(* IEC 61131-3 sources: daoli-st-library/DL_Motion (part 21) *)

(* ---- FB_DL_ZoneSpeedTrim.st ---- *)
(*==============================================================================
 * 组件名称 (Component)  : FB_DL_ZoneSpeedTrim
 * 所属子库 (Sublibrary) : DL_Motion
 * 当前版本 (Version)    : 1.0.0
 * 兼容性   (Platform)   : CODESYS 3.5+ / TwinCAT 3 / 汇川 InoProShop / 施耐德 Machine Expert
 *                         仅依赖 Standard.library（MIN / MAX / ABS），零厂商私有库
 * 功能描述 (Function)   : 轴位置区段差异化限速：按轴实际位置命中区段表（fStartMm/fEndMm/
 *                         fVmaxMmS）改写指令速度上限：命中 → fVCmd = MIN(fVout, fVmaxZone)；
 *                         表外 → MIN(fVout, fVDefault)。eCurZone 出当前命中区段号
 *                         （0=表外）。适用机械臂/桁架近人区、近件区、换向区差异化限速。
 * 接口     (Interface)  : 输入 fPosMm 轴实际位置（mm）、aZone 区段表（定长 1..nZoneMax）、
 *                         nZoneCount 有效区段数、fVDefaultMmS 表外默认限速（mm/s）、
 *                         fVoutMmS 当前指令速度（mm/s）、bReset 复位；输出 fVCmdMmS 限幅
 *                         后指令（mm/s）、eCurZone 当前命中区段号（0=表外）、bCapped
 *                         触限幅、bCfgBad 区段表非法（锁存）、bError 故障标志。
 * 边界     (Boundary)   : ① **属主边界（写死）：本件只做区段限速改写，不做静态软限位
 *                         报警、不接管轴使能**（静态软限位归 `FB_DL_SoftLimitGuard`）。
 *                         ② 区段表校验锁存 bCfgBad（表非法比静默错限速危险）：fStart>fEnd
 *                         （倒序）、fVmax<=0、任两区段重叠（含区间闭端相交）→ 锁存；
 *                         bCfgBad 期输出保守限速 MIN(fVout, fVDefault)，解除沿 =
 *                         bReset 上升沿。
 *                         ③ fStart<=fEnd 判据用浮点 < / > 比较，禁 = 判等（R28）。
 *                         ④ 表满 nZoneMax 钳位：nZoneCount > nZoneMax 按上限处理并置
 *                         组态当拍错。
 *                         ⑤ 非有限位置 → 冻结上次输出并置当拍 bError（R245）。
 *                         ⑥ 零全局耦合（无 GVL / VAR_EXTERNAL / 物理地址）。
 * 分工声明 (Scope)      : 与 `FB_DL_SoftLimitGuard` 分工：动态区段限速（本件）≠ 静态软
 *                         限位报警（那件）；与 `FB_DL_ConveyorZone` 分工：运动限速 ≠
 *                         输送段跟踪。
 * 来源标签 (Source Tag) : T1-6 ◐（PLCopen MC 语义只借限速语义，区段表结构自研）
 * 码表     (Codes)      : 本件不占用任何全局数字码位。出口为 LREAL 限速 + UDINT 区号 +
 *                         BOOL 组；数字码位待主控收口阶段统一派号。
 * 红线自检 (Redline)    : R1 ✓ 零 GVL/VAR_EXTERNAL ｜ R2 ✓ 零 %I/%Q/%M ｜ R3 ✓ 纯 IEC 61131-3
 *                         R4 ✓ 表校验锁存 + 浮点禁等 + 非有限冻结 + 表满钳位 ｜ R5 ✓ 声明逐行同行双语注释
 *                         R6 N/A（查表无状态机） ｜ R7 ✓ 一 R_TRIG 段 0 无条件刷新
 * 修订历史 (Revision)   : 2026-11-20  v1.0.0  R48 首版（批次 3 · 序号 15）
 *                         验收向量：命中区段按 fVmax 限幅；表外用默认值；倒序/重叠表 →
 *                         bCfgBad 锁存保守限速；nZoneCount 超上限钳位。
 *==============================================================================*)

TYPE ST_DL_ZoneSpeed :
STRUCT
    fStartMm  : LREAL;   // 区段起点（含端点） [mm] / Zone start, inclusive [mm]
    fEndMm    : LREAL;   // 区段终点（含端点） [mm] / Zone end, inclusive [mm]
    fVmaxMmS  : LREAL;   // 区段速度上限，域 > 0 [mm/s] / Zone speed ceiling [mm/s]
END_STRUCT
END_TYPE

FUNCTION_BLOCK FB_DL_ZoneSpeedTrim
VAR_INPUT
    fPosMm      : LREAL := 0.0;   // 轴实际位置 [mm] / Axis actual position [mm]
    aZone       : ARRAY[1..8] OF ST_DL_ZoneSpeed;   // 区段表（定长，nZoneCount 指明有效前段） / Zone table, fixed length
    nZoneCount  : UDINT := 0;     // 有效区段数（0=全表外） [段] / Valid zone count
    fVDefaultMmS: LREAL := 500.0; // 表外默认限速，域 > 0 [mm/s] / Default speed ceiling outside table [mm/s]
    fVoutMmS    : LREAL := 0.0;   // 当前指令速度（限幅前） [mm/s] / Command speed before capping [mm/s]
    bReset      : BOOL := FALSE;  // 复位，上升沿清 bCfgBad 锁存 [-] / Reset, rising edge clears cfg latch
END_VAR
VAR_OUTPUT
    fVCmdMmS : LREAL;            // 限幅后指令速度 [mm/s] / Capped command speed [mm/s]
    eCurZone : UDINT;            // 当前命中区段号（1..n，0=表外） [段] / Current zone number, 0 = outside
    bCapped  : BOOL;             // 本拍触限幅（fVCmd < fVout） [-] / Capped this scan
    bCfgBad  : BOOL;             // 区段表非法（锁存） [-] / Illegal zone table, latched
    bError   : BOOL;             // 故障标志（组态锁存 ∨ 非有限当拍） [-] / Error flag
END_VAR
VAR
    _nCount  : DINT;             // 钳位后有效区段数 [段] / Clamped valid zone count
    _nHit    : DINT;             // 命中区段号（0=表外） [段] / Hit zone number
    _fCap    : LREAL;            // 当拍生效速度上限 [mm/s] / Effective speed ceiling
    _fVCmd   : LREAL := 0.0;     // 输出锁存镜像（非有限冻结源） / Output latch mirror
    _bCfgLatch: BOOL;            // 表非法锁存位（解除沿 = bReset 上升沿） / Latched table fault
    _bErrScan: BOOL;             // 当拍错误内部量（钳位超限/非有限） / Per-scan error internal
    _bNonFin : BOOL;             // 位置非有限当拍量 [-] / Non-finite position this scan
    i        : DINT;             // 区段循环索引 / Zone loop index
    j        : DINT;             // 重叠校验内层索引 / Overlap check inner index
    rtReset  : R_TRIG;           // 复位沿实例，段 0 无条件调用 / Reset edge instance
END_VAR
VAR CONSTANT
    DL_ZST_NMAX : DINT  := 8;        // 区段表定长上限 [段] / Zone table length ceiling
    DL_ZST_EPS  : LREAL := 0.0;      // 非有限差值判零基准 [-] / Non-finite difference zero base
END_VAR

(* —— 段 0：非有限判 + 表满钳位 + 沿刷新 —— *)
_bNonFin := (fPosMm <> fPosMm) OR ((fPosMm - fPosMm) <> DL_ZST_EPS);   // 位置非有限（R245） / Non-finite position
_nCount := UDINT_TO_DINT(nZoneCount);        // 区段数转 DINT（UDINT 超界由下步钳位） / Convert count
IF _nCount > DL_ZST_NMAX THEN
    _nCount := DL_ZST_NMAX;                  // 表满钳位（头注释④） / Clamp to table ceiling
    _bErrScan := TRUE;                       // 超限置当拍组态错 / Mark per-scan error
END_IF
IF _nCount < 0 THEN
    _nCount := 0;                            // UDINT 溢出到 DINT 负值兜底 / Overflow fallback to zero
    _bErrScan := TRUE;                       // 记当拍错 / Mark per-scan error
END_IF
IF fVDefaultMmS <= 0.0 THEN
    _bErrScan := TRUE;                       // 默认限速组态闸（当拍报） / Default ceiling gate
END_IF
rtReset(CLK := bReset);                      // 复位沿，每拍必调 / Reset edge, every scan

(* —— 段 1：复位沿 —— *)
IF rtReset.Q THEN
    _bCfgLatch := FALSE;                     // 清表非法锁存 / Clear table latch
END_IF

(* —— 段 2：区段表校验（倒序 / 非正限速 / 重叠 → 锁存） —— *)
IF NOT _bCfgLatch THEN
    FOR i := 1 TO _nCount DO
        IF (aZone[i].fStartMm > aZone[i].fEndMm) OR (aZone[i].fVmaxMmS <= 0.0) THEN
            _bCfgLatch := TRUE;              // 倒序或非正限速：表非法锁存（头注释②） / Reversed or bad ceiling: latch
        END_IF
    END_FOR
    FOR i := 1 TO _nCount DO
        FOR j := (i + 1) TO _nCount DO
            IF (aZone[j].fStartMm <= aZone[i].fEndMm) AND (aZone[i].fStartMm <= aZone[j].fEndMm) THEN
                _bCfgLatch := TRUE;          // 任两区段闭区间相交：重叠非法锁存 / Overlapping zones: latch
            END_IF
        END_FOR
    END_FOR
END_IF

(* —— 段 3：限速主算（表非法期保守限速；非有限冻结） —— *)
_nHit := 0;                                  // 命中区号预清 / Hit preset
_fCap := fVDefaultMmS;                       // 上限预置默认值 / Preset default ceiling
IF (NOT _bCfgLatch) AND (NOT _bNonFin) AND (NOT _bErrScan) THEN
    FOR i := 1 TO _nCount DO
        IF (fPosMm >= aZone[i].fStartMm) AND (fPosMm <= aZone[i].fEndMm) THEN
            _nHit := i;                      // 位置命中区段（闭区间含端点，浮点仅用 < > 比较） / Position hits zone
            _fCap := aZone[i].fVmaxMmS;      // 区段限速生效 / Zone ceiling effective
        END_IF
    END_FOR
    _fVCmd := fVoutMmS;                      // 基准指令速度 / Base command speed
    IF _fVCmd > _fCap THEN
        _fVCmd := _fCap;                     // 超区段限速：限幅 / Cap to zone ceiling
    END_IF
ELSIF _bCfgLatch OR _bErrScan THEN
    _fVCmd := fVoutMmS;                      // 组态病期从默认保守限速出发 / Config fault: conservative base
    IF _fVCmd > fVDefaultMmS THEN
        _fVCmd := fVDefaultMmS;              // 保守限幅到表外默认值 / Conservative cap
    END_IF
END_IF
(* 非有限位置分支：无赋值 → _fVCmd 冻结上次值（头注释⑤） *)

(* —— 段 4：出口单点映射（名实双出口同源，R191） —— *)
fVCmdMmS := _fVCmd;                          // 限速输出 / Capped speed outlet
eCurZone := DINT_TO_UDINT(_nHit);            // 命中区号出口（0=表外） / Zone number outlet
bCapped  := _fVCmd < fVoutMmS;               // 触限幅判定（严格小于，浮点禁等兼容） / Capped flag
bCfgBad  := _bCfgLatch;                      // 表非法出口 / Table fault outlet
bError   := _bCfgLatch OR _bErrScan OR _bNonFin;   // 故障标志三源合一 / Error flag

END_FUNCTION_BLOCK

(* ---- FB_DL_AxisBrakeSeq.st ---- *)
(*
    FB_DL_AxisBrakeSeq —— 伺服抱闸时序
    ------------------------------------------------------------------
    分类      : DL_Motion / AxisSafety
    前缀      : FB_DL_
    版本      : 1.0.1
    溯源      : T1-6 PLCopen（只借「使能 / 抱闸属于轴生命周期授权动作」的公开语义，
                MC_Power 类功能块的使能时序纪律）；T2-4 S7 Motion 抱闸组织为次源；
                两序状态机、超时取舍、码位 100% 自有；clean-room 重写，
                未复制任何闭源厂商源码，参考实现仅限 MIT/Apache 许可
    道莅 clean-room 防御性实现：语义借鉴、代码与码位 100% 自有
    平台      : 纯 IEC 61131-3，CODESYS V3.5+ / TwinCAT 3 / InoProShop / Machine Expert 通用
    作者      : 道莅代码库 · PLC编程专家（R22 批 4 · #12）
    ------------------------------------------------------------------
    功能说明  : 伺服轴「上电」与「断电」两条机械-电气强制顺序的唯一屬主件。
                本件只输出两个有序命令（抱闸释放命令、伺服使能命令），
                不发运动指令、不自造轴状态枚举，轴状态唯一属主仍在轴功能块。
    两条序（顺序写反即掉轴，此处文字画时序，编码与之一一对应）:
                上电序 A：bEnableReq↑
                          → bBrakeReleaseCmd := TRUE
                          → 等「抱闸释放到位」（有反馈等反馈；无反馈等 tBrakeRelease）
                          → bServoEnable := TRUE
                          → eEnabled
                  理由：先使能后释放，电机顶着抱闸出力，抱闸片烧蚀。
                断电序 B：bEnableReq↓
                          → eStopping：保持带使能、保持抱闸打开
                          → 等 |fActVel| < fStandstillVel 连续 tStandstill
                          → bBrakeReleaseCmd := FALSE（抱闸闭合）
                          → 等 tBrakeHold（机械闭合建立力矩）
                          → bServoEnable := FALSE
                          → eDisabled
                  理由：先断使能后抱闸，轴在自由态下滑落；抱闸未建立力矩就断使能同样滑落。
    设计取舍  : ① 断电序中轴未在 tFbTimeout 内静止 → 报 02EB 并「拒绝断使能」：
                   保持带使能 + 保持抱闸打开，把轴钉在原位。宁可报警停线，不可掉轴。
                   若此时伺服本就没有使能（无转矩可用），则无「拒绝」可言，
                   改为立即闭合抱闸并报警——无转矩时抱闸是唯一能拦住轴的机构，
                   宁可磨损抱闸片也不让它自由滑落。两条支路靠 _bServoOn 上一拍快照区分。
                ② 抱闸释放反馈超时 → 报 02EA 并「禁止使能」，直接全失电
                   （弹簧制动器失电即抱死，是唯一安全侧）。
                ③ 无反馈现场（bBrakeFbAvailable = FALSE）按纯时间序列放行，
                   报信息 01D5；该风险由现场调试承担，头注释即为此留档。
    错误码    : 16#0004_01D5 无抱闸释放反馈，已按纯时间序列放行——信息级，正常防御
                16#0004_01D6 等待延长后放行（抱闸释放反馈迟到但收到 / 断电序静止窗因
                              速度抖动反复重启已延长等待）——信息级，两处共用本码，
                              靠所处状态区分，不得据此拒绝动作（R90）
                16#0004_02EA 抱闸释放反馈超 tFbTimeout，禁止使能——故障级，全失电
                16#0004_02EB 断电序轴未静止超 tFbTimeout，拒绝断使能——故障级，
                             有转矩时保持带使能 + 抱闸打开
                16#0004_02EC 序列参数非法 / 采样非有限 / 状态机落 ELSE 兜底——故障级
                             （三支复用，R90；靠进入路径区分，均回 eFault 并全失电）
    码位总账  : 16#0004_01D5 用 / 16#0004_01D6 用 ｜ 16#0004_02EA 用 / 16#0004_02EB 用 / 16#0004_02EC 用
    状态机    : E_DL_BrakeSeqState（eIdle / eReleasing / eEnabled / eStopping / eBraking
                / eDisabled / eFault），CASE 含 ELSE 兜底，ELSE 置 16#0004_02EC 并回 eFault；
                失能请求无条件经 eStopping，eEnabled 不得直跳 eDisabled（R71）。
    采样约定  : 五个 TON 实例在本体最前部无条件调用（R40），每段一只实例、绝不跨段复用；
                段转出统一走「断输入一拍」标志（_bRelBreak / _bStopBreak / _bHoldBreak），
                断一拍标志在对应 TON 调用之后立刻自清，避免下一拍再吞掉计时。
                本件不读系统时钟，时间全部来自 TIME 引脚。
    依赖      : 仅 Standard.library（TON / ABS / MIN / MAX / LIMIT），
                不引用任何其他 DL_ 子库（DL_Motion/VERSION.md 硬约束）。
    验收向量  :
                V1 域外早退：fStandstillVel = 0 → 02EC、bError=TRUE、bValid=FALSE、
                   两命令全 FALSE（弹簧制动器失电抱死）。
                V2 上限截断/超时：bBrakeReleaseFb 恒 FALSE 且 bBrakeFbAvailable=TRUE
                   → tFbTimeout 到 → 02EA、bServoEnable 恒 FALSE、bBrakeReleaseCmd 转 FALSE。
                V3 跨段时序：eEnabled 中 bEnableReq↓ 同拍 fActVel = 50 mm/s（未静止）
                   → 先入 eStopping 且 bServoEnable 保持 TRUE、bBrakeReleaseCmd 保持 TRUE，
                   tFbTimeout 后才报 02EB；不得同拍闭合抱闸。
                V4 恢复/复位首拍：抱闸闭合后立即 bEnableReq↑（eBraking 期间）
                   → 不得半途重启上电序，须走完 eBraking → eDisabled → eIdle → eReleasing。
    红线自检  : 1 全局变量声明零使用 / 外部变量访问零使用 / 物理地址零使用 —— 通过，全部量经引脚注入
                2 纯 IEC 61131-3 跨平台 —— 通过，仅 Standard.library
                3 防御性编程 —— 通过，浮点判等全用绝对值阈、无非有限值穿透、无除法
                4 声明行同行中英双语注释 + 单位 —— 通过，逐行附注（含枚举成员）
                5 ENUM + CASE 且含 ELSE 兜底 —— 通过，两条 CASE（主状态机 / 输出映射）
                6 TON / R_TRIG 无条件刷新 —— 通过，段 1 全部实例先行调用
                7 无魔法数 —— 通过，阈值与时间全部为引脚或 VAR CONSTANT
    修订记录  : 2026-11-16 v1.0.0 首次入库（R22 批 4 · #12）
                2026-11-16 v1.0.1 R22 终审勘误：tBrakeRelease 引脚注释原写「有反馈时
                作为最短等待」，实现实际为「反馈到达即采信」，注释对齐实现（不改时序
                代码）；并显式声明配置约束 tFbTimeout > tBrakeRelease——超时窗
                （fbRelFeedback）与标称等待（fbRelease）同拍起算，若超时窗不大于
                标称等待，会在标称时间之前误报 02EA
*)
TYPE E_DL_BrakeSeqState :
(
    eIdle      := 0,     // 待机，两命令全失电，等使能请求上升沿 / idle, both commands de-energised, waiting for the enable request
    eReleasing := 10,    // 抱闸释放中，等释放到位或时间放行，伺服仍未使能 / releasing the brake, servo not yet enabled
    eEnabled   := 20,    // 已使能，抱闸打开且伺服带转矩，可接受运动指令 / enabled, brake open and servo energised
    eStopping  := 30,    // 断电序等待静止，保持带使能 + 保持抱闸打开 / stopping, waiting for standstill while keeping enable and brake open
    eBraking   := 40,    // 抱闸已闭合，等 tBrakeHold 建立机械力矩 / brake engaged, waiting for the mechanical torque build-up
    eDisabled  := 50,    // 已失电，抱闸闭合，伺服失能，可接受新使能请求 / disabled, brake engaged and servo de-energised
    eFault     := 60     // 故障，出口按 _bHoldEnableOnFault 决定保持或全失电 / fault, outputs follow the hold flag
);
END_TYPE

FUNCTION_BLOCK FB_DL_AxisBrakeSeq
VAR_INPUT
    bEnableReq        : BOOL;                  // 使能请求（上升沿启动上电序，下降沿启动断电序）/ enable request, rising edge starts the power-up sequence
    fActVel           : REAL;                  // 轴实际速度 [mm/s]，取绝对值参与静止判定 / axis actual velocity [mm/s], absolute value used for the standstill test
    fStandstillVel    : REAL := 1.0;           // 静止判定速度阈 [mm/s]，必须大于 0 / standstill velocity threshold [mm/s], must exceed zero
    bBrakeReleaseFb   : BOOL;                  // 抱闸释放到位反馈，TRUE = 已释放 / brake released feedback, TRUE = fully released
    bBrakeFbAvailable : BOOL := TRUE;          // FALSE 时按纯时间序列（无反馈现场）/ FALSE = time-based sequence only on a site without feedback
    tBrakeRelease     : TIME := T#200MS;       // 抱闸释放标称等待 [ms]，无反馈时按此放行；有反馈时反馈到达即采信（不做最短等待）；超时窗自进相起算，须配置 tFbTimeout > tBrakeRelease / brake release nominal wait [ms]; without feedback the release is time-based, with feedback the acknowledgement is trusted on arrival (no minimum wait); the timeout window starts at phase entry, so tFbTimeout must exceed this value
    tBrakeHold        : TIME := T#300MS;       // 抱闸闭合保持等待 [ms]，建立机械力矩 / brake hold wait [ms] for the mechanical torque build-up
    tStandstill       : TIME := T#100MS;       // 静止确认时间 [ms]，必须大于 0 / standstill confirmation time [ms], must exceed zero
    tFbTimeout        : TIME := T#2S;          // 序列超时 [ms]，必须大于 0 / sequence timeout [ms], must exceed zero
END_VAR
VAR_OUTPUT
    bServoEnable      : BOOL;                  // 伺服使能命令，上电序最后置位、断电序最先复位 / servo enable command, set last on power-up and cleared first on power-down
    bBrakeReleaseCmd  : BOOL;                  // 抱闸释放命令，上电序最先置位、断电序先于使能复位 / brake release command, set first on power-up and cleared before the enable drops
    bSeqDone          : BOOL;                  // 断电序完成单拍脉冲，发布后即刻自清 / one-scan pulse at power-down completion, self-cleared right after publishing
    eErr              : UDINT;                 // 错误码，0 表示无错 / error code, 0 means no error
    bError            : BOOL;                  // 故障级标志，仅故障级错误置位 / fault-class flag, set only on fault-level codes
    bValid            : BOOL;                  // 输出可用标志，= NOT bError / outputs valid flag, equals NOT bError
END_VAR
VAR
    fbRelease         : TON;                   // 抱闸释放最短等待定时器，仅 eReleasing 使用 / brake release minimum wait, used in eReleasing only
    fbRelFeedback     : TON;                   // 抱闸释放反馈超时定时器，仅 eReleasing 使用 / release feedback timeout, used in eReleasing only
    fbStandstill      : TON;                   // 静止确认定时器，仅 eStopping 使用 / standstill confirmation timer, used in eStopping only
    fbStopTimeout     : TON;                   // 断电序总超时定时器，仅 eStopping 使用 / power-down timeout, used in eStopping only
    fbBrakeHold       : TON;                   // 抱闸闭合保持定时器，仅 eBraking 使用 / brake hold timer, used in eBraking only
    _bRelBreak        : BOOL;                  // eReleasing 两只定时器的断输入一拍标志 / break-input flag for the two timers of eReleasing
    _bStopBreak       : BOOL;                  // eStopping 两只定时器的断输入一拍标志 / break-input flag for the two timers of eStopping
    _bHoldBreak       : BOOL;                  // eBraking 定时器的断输入一拍标志 / break-input flag for the timer of eBraking
    _bServoOn         : BOOL;                  // 上一拍伺服使能快照，断电序与故障出口用 / previous-scan servo enable snapshot used by the stop phase and the fault exit
    _bStill           : BOOL;                  // 本拍静止条件（速度绝对值小于阈）/ standstill condition of this scan
    _bStillPrev       : BOOL;                  // 上一拍静止条件，用于捕捉稳定窗重启 / previous-scan standstill condition, catches a restarted window
    _bStopExtend      : BOOL;                  // 断电序等待被延长标志（稳定窗重启过一次）/ stop-phase wait extension flag, set once per sequence
    _bRelLate         : BOOL;                  // 抱闸释放反馈迟到标志，按序只报一次 / late release feedback flag, reported once per sequence
    _bFsmBad          : BOOL;                  // 采样非有限或参数非法标志，供码位链使用 / non-finite sample or illegal parameter flag feeding the code chain
    _bHoldEnableOnFault : BOOL;                // 故障出口「保持带使能 + 抱闸打开」锁存开关，仅 02EB 且有转矩时置位，离开故障态才清 / latched fault-exit hold switch, set only by 02EB when the drive had torque and cleared when leaving the fault state
    _uErrLatch        : UDINT;                 // 故障码锁存副本，故障态每拍重发布，防止段 2 预置冲掉 / latched fault code republished every scan inside the fault state
    _bDonePulse       : BOOL;                  // 断电序完成脉冲源，段 2 发布后立刻自清 / completion pulse source, published then cleared in segment 2
    _eState           : E_DL_BrakeSeqState;    // 当前状态 / current state
END_VAR
VAR CONSTANT
    DL_BS_INF_GUARD : REAL := 4.0E38;          // 非有限幅值判定阈值（大于 REAL 最大值）[mm/s] / non-finite magnitude guard above the REAL maximum [mm/s]
    DL_BS_ZERO      : REAL := 0.0;             // 零值常量，避免裸字面量 [无量纲] / zero constant, avoids a bare literal [dimensionless]
    DL_BS_T_ZERO    : TIME := T#0S;            // 零时间常量，用于参数门禁 / zero time constant used by the parameter gate
END_VAR

// 段 1｜五个 TON 无条件周期刷新（红线 6：严禁放入 IF / CASE，也严禁跨段复用实例）
// segment 1, five TON instances refreshed unconditionally, one instance per segment and never shared
fbRelease(IN := (_eState = E_DL_BrakeSeqState.eReleasing) AND (NOT _bRelBreak), PT := tBrakeRelease);
fbRelFeedback(IN := (_eState = E_DL_BrakeSeqState.eReleasing) AND (NOT _bRelBreak), PT := tFbTimeout);
_bRelBreak := FALSE;                            // 断输入标志用后即刻自清，避免下一拍再吞计时 / the break flag clears right after the call so the next scan times normally
_bStill := ABS(fActVel) < fStandstillVel;       // 本拍静止条件，绝对速度与阈比较 / standstill condition of this scan
fbStandstill(IN := (_eState = E_DL_BrakeSeqState.eStopping) AND (NOT _bStopBreak) AND _bStill, PT := tStandstill);
fbStopTimeout(IN := (_eState = E_DL_BrakeSeqState.eStopping) AND (NOT _bStopBreak), PT := tFbTimeout);
_bStopBreak := FALSE;                           // 断输入标志用后即刻自清 / the break flag clears right after the call
fbBrakeHold(IN := (_eState = E_DL_BrakeSeqState.eBraking) AND (NOT _bHoldBreak), PT := tBrakeHold);
_bHoldBreak := FALSE;                           // 断输入标志用后即刻自清 / the break flag clears right after the call

// 段 2｜输出与错误状态预置（单拍标志在此发布后立刻自清，R25 三律）
// segment 2, preset outputs and error status; the one-scan flag is published and cleared here
eErr := 0;                                      // 预置无错误 / preset no error
bError := FALSE;                                // 预置无故障标志 / preset no error flag
bSeqDone := _bDonePulse;                        // 发布上一拍置的完成脉冲 / publish the completion pulse latched last scan
_bDonePulse := FALSE;                           // 发布即自清，保证只出现一拍 / clear right after publishing so the pulse lasts exactly one scan

// 故障态的错误码与保持开关是锁存量：每拍从锁存副本重新发布，绝不因本段预置被冲掉（R45）
// inside the fault state the code and the hold switch are latched values republished every scan, the preset above cannot erase them
IF _eState = E_DL_BrakeSeqState.eFault THEN
    eErr := _uErrLatch;                         // 重发布锁存故障码，HMI 不会看到码位闪断 / republish the latched code so the HMI never sees it drop out
    bError := TRUE;                             // 故障态恒置故障标志 / the fault flag stays raised inside the fault state
END_IF

// 段 3｜参数与采样门禁：任一非法即全失电并锁死在本拍，不进状态机
// segment 3, parameter and sample gate; any violation de-energises at once and skips the state machine
IF (fStandstillVel <= DL_BS_ZERO)
   OR (tStandstill <= DL_BS_T_ZERO)
   OR (tFbTimeout <= DL_BS_T_ZERO) THEN
    _bFsmBad := TRUE;                           // 静止阈非正 / 确认时间为零 / 超时为零，序列无从判定 / the standstill threshold or a duration is not positive
ELSE
    _bFsmBad := FALSE;                          // 参数合法 / parameters are legal
END_IF

// 非有限采样检测：NaN 用自不自等捕获，±Inf 用幅值门捕获（REAL 最大约 3.4E38）
// non-finite sample detection, NaN via self-inequality and plus/minus infinity via the magnitude guard
IF (fActVel - fActVel) <> (fActVel - fActVel) THEN
    _bFsmBad := TRUE;                           // NaN / not a number
ELSIF ABS(fActVel) > DL_BS_INF_GUARD THEN
    _bFsmBad := TRUE;                           // ±Inf / plus or minus infinity
END_IF

IF _bFsmBad THEN
    eErr := 16#0004_02EC;                       // 故障级：参数非法或采样非有限（与兜底复用，R90）/ fault: illegal parameter or non-finite sample, shared with the fallback
    bError := TRUE;                             // 置故障标志 / raise the fault flag
    _uErrLatch := 16#0004_02EC;                 // 锁存故障码，故障态整段可观测 / latch the code so it stays observable for the whole fault state
    _bHoldEnableOnFault := FALSE;               // 参数不可信时全失电，弹簧制动器抱死 / de-energise when the parameters cannot be trusted, the spring brake locks
    _bRelBreak := TRUE;                         // 三组定时器全部断输入重启 / restart every timer group
    _bStopBreak := TRUE;
    _bHoldBreak := TRUE;
    _bServoOn := FALSE;                         // 快照清零，防止故障出口误保持 / clear the snapshot so the fault exit cannot hold by accident
    _eState := E_DL_BrakeSeqState.eFault;       // 转故障 / go to fault
END_IF

// 段 4｜等待延长观测（信息 01D6 的两处触发源，按序各报一次）
// segment 4, wait-extension observation, the two triggers of information code 01D6, once per sequence each
IF (_eState <> E_DL_BrakeSeqState.eReleasing) AND (_eState <> E_DL_BrakeSeqState.eStopping) THEN
    _bRelLate := FALSE;                         // 离开两序即清迟到标志，下一序可再报 / clear the late flag outside both phases so the next sequence can report again
    _bStopExtend := FALSE;                      // 清断电序延长标志 / clear stop-phase extension flag
END_IF

IF (_eState = E_DL_BrakeSeqState.eStopping) AND _bStillPrev AND (NOT _bStill) THEN
    _bStopExtend := TRUE;                       // 静止窗被打断，本轮等待将被延长 / the standstill window was interrupted, this stop will take longer
END_IF
_bStillPrev := _bStill;                         // 更新上一拍静止条件 / update the previous-scan standstill condition

// 段 5｜主状态机：两条序逐态编码，顺序即安全（R71：eEnabled 不得直跳 eDisabled）
// segment 5, the main state machine; the two sequences are encoded state by state and the order itself is the safety measure
CASE _eState OF
E_DL_BrakeSeqState.eIdle:
    // 待机：全失电，只在使能请求为真时启动上电序 A / idle, everything de-energised, start sequence A only when the request is present
    IF bEnableReq AND (NOT _bFsmBad) THEN
        _bRelBreak := TRUE;                     // 释放等待定时器断一拍重启 / restart the release timers with one scan of FALSE input
        _eState := E_DL_BrakeSeqState.eReleasing;   // 进释放相，下一拍输出段置抱闸释放命令 / enter the release phase, the output map asserts the release command next scan
    END_IF

E_DL_BrakeSeqState.eReleasing:
    // 上电序 A 第 2 步：等抱闸释放到位（有反馈等反馈，无反馈等时间放行）
    // power-up step 2, wait for the brake release, either the feedback or the time-based release
    IF bBrakeFbAvailable THEN
        IF fbRelease.Q AND (NOT bBrakeReleaseFb) THEN
            _bRelLate := TRUE;                  // 标称时间到但反馈未到，转为延长等待 / the nominal time elapsed without feedback, switch to an extended wait
        END_IF
        IF bBrakeReleaseFb THEN
            IF _bRelLate THEN
                eErr := 16#0004_01D6;           // 信息级：反馈迟到但已收到，按延长等待放行 / info: the feedback arrived late and the extended wait released it
            END_IF
            _eState := E_DL_BrakeSeqState.eEnabled;     // 释放到位，允许使能 / the brake is released, enabling is allowed
        ELSIF fbRelFeedback.Q THEN
            eErr := 16#0004_02EA;               // 故障级：释放反馈超时，禁止使能 / fault: release feedback timeout, enabling is forbidden
            bError := TRUE;                     // 置故障标志 / raise the fault flag
            _uErrLatch := 16#0004_02EA;         // 锁存故障码 / latch the code
            _bHoldEnableOnFault := FALSE;       // 全失电，抱闸抱死 / de-energise so the spring brake locks
            _eState := E_DL_BrakeSeqState.eFault;
        END_IF
    ELSE
        IF fbRelease.Q THEN
            _eState := E_DL_BrakeSeqState.eEnabled;     // 无反馈现场：时间到即放行 / no feedback on site, the elapsed time releases it
            eErr := 16#0004_01D5;               // 信息级：无反馈按纯时间序列（风险由现场调试承担）/ info: time-based sequence without feedback, the risk is borne on site
        END_IF
    END_IF
    // 上电序被撤回：不得半途使能，转断电序收尾（抱闸仍打开，先等静止再闭合）
    // the power-up request was withdrawn, never enable halfway and fall through to the stop phase
    IF NOT bEnableReq THEN
        _bStopBreak := TRUE;                    // 静止与超时定时器断一拍重启 / restart the standstill and timeout timers
        _eState := E_DL_BrakeSeqState.eStopping;
    END_IF

E_DL_BrakeSeqState.eEnabled:
    // 已使能：抱闸打开 + 伺服带转矩，断电请求落下即进断电序 B，绝不经由任何捷径
    // enabled, brake open and servo energised; a falling request enters sequence B and never takes a shortcut
    IF NOT bEnableReq THEN
        _bStopBreak := TRUE;                    // 静止与超时定时器断一拍重启 / restart the standstill and timeout timers
        _eState := E_DL_BrakeSeqState.eStopping;    // 必须经 eStopping（R71）/ must pass through eStopping
    END_IF

E_DL_BrakeSeqState.eStopping:
    // 断电序 B 第 1 步：等静止。此处只判不动，抱闸保持打开、使能保持
    // power-down step 1, wait for standstill; nothing moves here, the brake stays open and the enable is held
    IF fbStandstill.Q THEN
        _bHoldBreak := TRUE;                    // 抱闸保持定时器断一拍重启 / restart the brake hold timer
        _eState := E_DL_BrakeSeqState.eBraking;// 静止确认，允许闭合抱闸 / standstill confirmed, the brake may now engage
        IF _bStopExtend THEN
            eErr := 16#0004_01D6;               // 信息级：静止确认窗被抖动打断，等待已延长 / info: the standstill window was interrupted, the wait was extended
        END_IF
    ELSIF fbStopTimeout.Q THEN
        eErr := 16#0004_02EB;                   // 故障级：轴未静止超时 / fault: the axis did not reach standstill in time
        bError := TRUE;                         // 置故障标志 / raise the fault flag
        _uErrLatch := 16#0004_02EB;             // 锁存故障码 / latch the code
        _bHoldEnableOnFault := _bServoOn;       // 有转矩才拒绝断使能；无转矩时改由抱闸拦轴 / only hold the enable when the drive had torque, otherwise let the brake catch the axis
        _eState := E_DL_BrakeSeqState.eFault;
    END_IF
    // 断电序中使能请求又来了：先把本次断电序走完，不允许反向插入（V4 向量）
    // the request came back during the stop phase, finish the stop first and never insert a reverse step

E_DL_BrakeSeqState.eBraking:
    // 断电序 B 第 2 步：抱闸已闭合，等 tBrakeHold 建立机械力矩后才允许断使能
    // power-down step 2, the brake is engaged and the enable must survive the whole hold time
    IF fbBrakeHold.Q THEN
        _bDonePulse := TRUE;                    // 断电序完成脉冲，段 2 下一拍发布并自清 / latch the completion pulse, published and cleared by segment 2 next scan
        _eState := E_DL_BrakeSeqState.eDisabled;
    END_IF

E_DL_BrakeSeqState.eDisabled:
    // 已失电：全输出为假，接受新使能请求（请求仍在则一拍后重启上电序）
    // disabled, every output is false and a new request re-enters the power-up sequence one scan later
    IF bEnableReq AND (NOT _bFsmBad) THEN
        _eState := E_DL_BrakeSeqState.eIdle;    // 回待机，由待机态统一启动，避免两条启动路径 / return to idle so that a single start path exists
    END_IF

E_DL_BrakeSeqState.eFault:
    // 故障：只允许在请求已撤且参数已修好后复位；出口由输出映射段按 _bHoldEnableOnFault 决定
    // fault, reset is accepted only after the request is withdrawn and the parameters are repaired
    IF (NOT bEnableReq) AND (NOT _bFsmBad) THEN
        _bRelBreak := TRUE;                     // 三组定时器全部断输入重启 / restart every timer group
        _bStopBreak := TRUE;
        _bHoldBreak := TRUE;
        _eState := E_DL_BrakeSeqState.eIdle;    // 回待机 / return to idle
    END_IF

ELSE
    // 非法状态兜底：绝不静默停在未知态 / illegal state fallback, never stay silently in an unknown state
    eErr := 16#0004_02EC;                       // 故障级：状态机落 ELSE（与参数门禁复用，R90）/ fault: the state machine fell into ELSE, shared with the parameter gate
    bError := TRUE;                             // 置故障标志 / raise the fault flag
    _uErrLatch := 16#0004_02EC;                 // 锁存故障码 / latch the code
    _bHoldEnableOnFault := FALSE;               // 未知态一律全失电 / an unknown state always de-energises
    _bRelBreak := TRUE;                         // 三组定时器全部断输入重启 / restart every timer group
    _bStopBreak := TRUE;
    _bHoldBreak := TRUE;
    _eState := E_DL_BrakeSeqState.eFault;       // 回故障态 / go to fault
END_CASE

// 段 6｜输出映射（R72 双路径：段首已全部置假，此处按状态逐项置真，绝不漏项）
// segment 6, output map; the double-path rule presets everything to false first and asserts per state here
CASE _eState OF
E_DL_BrakeSeqState.eIdle:
    ;                                           // 待机：两命令保持假（弹簧制动器抱死）/ idle, both commands stay false and the spring brake holds
E_DL_BrakeSeqState.eReleasing:
    bBrakeReleaseCmd := TRUE;                   // 释放相：只给抱闸释放命令，伺服仍未使能 / release phase, only the brake release command, the servo is not enabled yet
E_DL_BrakeSeqState.eEnabled:
    bBrakeReleaseCmd := TRUE;                   // 已使能：抱闸打开 / enabled, the brake stays open
    bServoEnable := TRUE;                       // 已使能：伺服带转矩 / enabled, the servo is energised
E_DL_BrakeSeqState.eStopping:
    bBrakeReleaseCmd := TRUE;                   // 断电序：静止前抱闸必须保持打开 / stop phase, the brake must stay open until standstill
    bServoEnable := _bServoOn;                  // 断电序：保持上一拍使能，绝不提前断 / stop phase, hold the previous-scan enable and never drop it early
E_DL_BrakeSeqState.eBraking:
    bBrakeReleaseCmd := FALSE;                  // 抱闸闭合：命令已撤，机械抱死 / the brake engages because the release command is withdrawn
    bServoEnable := _bServoOn;                  // 保使能直到 tBrakeHold 走完 / keep the enable until the hold time elapses
E_DL_BrakeSeqState.eDisabled:
    ;                                           // 已失电：两命令保持假 / disabled, both commands stay false
E_DL_BrakeSeqState.eFault:
    bBrakeReleaseCmd := _bHoldEnableOnFault;    // 有转矩的 02EB 保持抱闸打开，其余全失电 / hold the brake open only for the torque case of 02EB
    bServoEnable := _bHoldEnableOnFault;        // 有转矩的 02EB 保持使能，其余全失电 / hold the enable only for that same case
ELSE
    ;                                           // 非法状态：两命令保持假，安全侧 / illegal state, both commands stay false, the safe side
END_CASE

// 段 7｜出口汇总：离开故障态即清锁存（保证下一次故障是全新判定），快照必须在输出映射之后更新
// segment 7, exit aggregation; leaving the fault state clears the latches and the snapshot follows the output map
IF _eState <> E_DL_BrakeSeqState.eFault THEN
    _uErrLatch := 0;                            // 清故障码锁存 / clear the latched fault code
    _bHoldEnableOnFault := FALSE;               // 清保持开关，故障出口默认全失电 / clear the hold switch, the fault exit defaults to full de-energisation
END_IF
_bServoOn := bServoEnable;                      // 上一拍伺服使能快照，供断电序与故障出口使用 / previous-scan enable snapshot used by the stop phase and the fault exit
bValid := NOT bError;                           // 输出可用 = 无故障级错误 / outputs are valid when no fault-level code is present
END_FUNCTION_BLOCK

(* ---- FB_DL_AxisHomingSeq.st ---- *)
(*==============================================================================
 * 组件名称 (Component)  : FB_DL_AxisHomingSeq
 * 所属子库 (Sublibrary) : DL_Motion
 * 当前版本 (Version)    : 1.0.1
 * 组件分类 (Category)   : 功能块（FUNCTION_BLOCK）· 轴回零序列状态机 · 工艺上层件
 * 兼容性   (Platform)   : CODESYS 3.5 / TwinCAT 3 / 汇川 InoProShop / Schneider
 *                         Machine Expert；仅依赖 Standard.library（TON / R_TRIG /
 *                         F_TRIG / MIN / MAX / ABS），零厂商方言
 * 接口依赖 (Depends)    : I_DL_MotionAxis / E_DL_AxisState（既有契约，Round 05）
 * 功能描述 (Function)   : 标准工业回零序列状态机。经轴接口引用驱动轴体，全部
 *                         序列动作由 MoveVelocity / Stop 组合出，本块绝不出任何
 *                         自有速度输出。四模式：限位开关回零 / 原点开关回零 /
 *                         Z 相脉冲精定位 / 扭矩堵转回零。慢速逼近-回退-再逼近-
 *                         标定时序。被动回零（外力移动轴监听参考事件）本轮不
 *                         实现，留矩阵扩产。
 * 设计要点 (Key notes)  : ① 双护栏：总超时（TON 自实现周期累积）+ 行程超限
 *                           （起点-当前位置绝对差 > fMaxTravel）；
 *                         ② 启动门禁：轴不在待机态 / 参数非法 / 可观测矛盾
 *                           （原点开关或所选限位启动时已压住）→ 拒绝并置
 *                           信息级 0004_0106；信号缺失类不可观测项（Z 相通道
 *                           无效、堵转阈值未组态）由调用方保证（头注释声明）；
 *                         ③ 标定职责边界：eCalibrate 仅完成受控停车与序列收口，
 *                           坐标系写入与轴回原标志置位由调用方联动 bDone 完成，
 *                           本块不直接写轴内部态（接口无位置写入域）；
 *                         ④ bTrack 中途插入 → 序列中止受控停车回空闲（R19）；
 *                         ⑤ R14：超时定时器 PT 变更显式断输入一拍使已计时归零。
 * 规格偏离留档 (R11)    : 规格引脚表未列回零方向，但四模式时序均需逼近方向
 *                         语义，补充 bDirNeg : BOOL 输入（TRUE=朝负方向回零）；
 *                         fMaxTravel 为规格正文明确的新增引脚（默认 1.0E6）。
 * 开源溯源 (Origin)     : 原创实现（参考 PLCopen Part 1-6 回零方式分类与西门子
 *                         Motion Control 对象语义，clean-room）。仅提取公开的
 *                         回零方式分类（限位/原点开关/Z 相/扭矩堵转）与
 *                         逼近-回退-再逼近-标定公开语义；实现与命名 100% 自有，
 *                         未参考任何厂商源码行。
 * 验收向量 (Acceptance) :
 *   V1 限位开关回零全链：逼近→限位上升沿→反向回退→限位下降沿→爬行再逼近→
 *      限位上升沿→标定→完成；V2 原点开关回零全链（逼近-回退-再逼近逐拍）；
 *   V3 Z 相精定位：爬行单向→Z 相上升沿→标定→完成；V4 堵转回零：爬行→
 *      堵转信号→标定→完成；V5 总超时 → 故障码 0004_0210；V6 行程超限 →
 *      0004_0211；V7 启动门禁（轴非待机/原点开关已压住）→ 信息级 0004_0106
 *      拒绝；V8 运行中途 bTrack → 受控停车回空闲（R19 必测）。
 * 故障码表 (Error codes):
 *   16#0004_0106【信息级】启动门禁/参数门禁拒绝（与 FB_DL_AxisRelativeMove
 *   同码同义，共用留档）；16#0004_0210【故障级】回零总超时；
 *   16#0004_0211【故障级】行程超限；16#0004_0212【故障级】中止/轴故障；
 *   16#0004_0213【故障级】序列指令被拒或非法状态兜底。
 * 修订历史 (Revision)   :
 *   2026-11-15  v1.0.0  首版入库（Round 06 · DL_Motion 回零/运动族）
 *   2026-11-15  v1.0.1  终审修复【严重】终态死锁：原实现 eDone/eAborted/
 *                       eFault 三态在 CASE 内无任何迁出路径，启动上升沿被
 *                       吞——首次回零完成后（或中止/故障后）永远无法再次
 *                       回零，仅 bTrack 可逃逸（R6 状态机跃迁完整性检查项
 *                       复现）。修法：新增段 5.5 终态重启借道逻辑——三终
 *                       态收到启动沿即回 eIdle，使同拍 eIdle 门禁分支受理
 *                       该沿（不吞沿、不要求双击）。引脚契约零变更。
 *============================================================================*)

(*-----------------------------------------------------------------------------
 * 调用示例 (Instance guide)：
 *   fbHome.iAxis := fbAxis;                       // 接口依赖注入
 *   fbHome(eMode := E_DL_HomingMode.eHomeSwitch,  // 周期调用
 *          bCmdStart := bStartHome, bDirNeg := TRUE,
 *          fHomingVel := 50.0, fCreepVel := 2.0, fAcc := 1000.0,
 *          fHomePosition := 0.0, tHomingTimeout := T#60S,
 *          bLimPos := swLimP, bLimNeg := swLimN, bHomeSw := swHome);
 *   IF fbHome.bDone THEN … 上层联动：写入轴坐标系 fHomePosition 并置轴回原标志（示例省略）
 *   注意：本块只驱动序列，坐标系建立由调用方在 bDone 后执行。
 *----------------------------------------------------------------------------*)

(*-----------------------------------------------------------------------------
 * 常见误用与现场提示 (Field notes)：
 *   1 启动时原点开关/所选限位已压住属可观测矛盾，本块拒绝启动（信息级
 *     0004_0106）；Z 相通道无效、堵转阈值未组态等不可观测项由调用方保证。
 *   2 eDone 态 bDone 保持 TRUE，回零完成后轴接口回原标志由上层联动；本块
 *     不重复标定，直到下一次 bCmdStart 上升沿。
 *   3 fHomePosition 在本块内不参与运算，作为标定值暂存引脚供上层读取写入
 *     轴坐标系（接口无位置写入域，职责边界见设计要点③）。
 *----------------------------------------------------------------------------*)

(*-----------------------------------------------------------------------------
 * 枚举: E_DL_HomingMode（归属 DL_Motion，与 FB_DL_AxisHomingSeq 同文件）
 * 含义: 回零方式选择。模式是组合矩阵而非厂商魔法数：本库仅取四种高频方式，
 *       取值不用任何厂商模式数值，其余方式留扩产。
 *----------------------------------------------------------------------------*)
{attribute 'strict'}
{attribute 'qualified_only'}
TYPE E_DL_HomingMode :
(
    eLimitSwitch := 1,   // 限位开关回零（Limit switch homing），以近端限位为参考
    eHomeSwitch  := 2,   // 原点开关回零（Home switch homing），独立原点开关
    eZeroPulse   := 3,   // Z 相脉冲精定位（Encoder zero pulse homing）
    eTorqueBlock := 4    // 扭矩堵转回零（Torque block homing），堵转阈值到达即原点
) UINT;
END_TYPE

(*-----------------------------------------------------------------------------
 * 枚举: E_DL_HomingStep（归属 DL_Motion，与 FB_DL_AxisHomingSeq 同文件）
 * 含义: 回零序列步。编号显式、间隔 10 预留扩展位，eFault 末位。
 *----------------------------------------------------------------------------*)
{attribute 'strict'}
{attribute 'qualified_only'}
TYPE E_DL_HomingStep :
(
    eIdle       := 0,    // 空闲：等待启动指令 / Idle: waiting for start command
    eApproach   := 10,   // 快速逼近（Z 相/堵转模式为爬行逼近）/ Fast approach (creep for zero-pulse/torque modes)
    eRetreat    := 20,   // 反向回退（限位模式全速回退/原点开关模式停车后爬行脱离）/ Reverse retreat
    eReapproach := 30,   // 爬行再逼近（Creep re-approach toward reference）
    eCalibrate  := 40,   // 标定原点（Calibrate home position），收口转受控停车
    eStopping   := 50,   // 受控停车等待停稳（Controlled stop, waiting standstill）
    eDone       := 60,   // 回零完成（Homing done），bDone 保持
    eAborted    := 70,   // 已中止（Aborted by command），受控停车后进入
    eFault      := 99    // 故障（Fault），仅重新启动可退出本块故障态
) UINT;
END_TYPE

FUNCTION_BLOCK FB_DL_AxisHomingSeq
VAR_INPUT
    eMode               : E_DL_HomingMode := E_DL_HomingMode.eHomeSwitch; // 回零模式（Homing mode），见 E_DL_HomingMode
    bCmdStart           : BOOL := FALSE;      // 回零启动（Homing start），上升沿生效
    bCmdAbort           : BOOL := FALSE;      // 回零中止（Homing abort），电平生效，触发受控停车
    bDirNeg             : BOOL := FALSE;      // 回零方向（Homing direction），TRUE=朝负方向逼近（规格外补充引脚，见头注 R11 留档）
    fHomingVel          : REAL := 50.0;       // 快速逼近速度（Homing approach velocity）[mm/s]，正值，默认 50.0
    fCreepVel           : REAL := 2.0;        // 爬行再逼近速度（Creep velocity）[mm/s]，正值，默认 2.0
    fAcc                : REAL := 1000.0;     // 回零加减速（Homing acceleration）[mm/s²]，正值，默认 1000.0
    fHomePosition       : REAL := 0.0;        // 标定原点位置值（Home position value）[mm]，暂存引脚，标定后由上层写入轴坐标系
    fMaxTravel          : REAL := 1.0E6;      // 行程护栏上限（Max travel guard）[mm]，|当前位置-起点| 超限即故障，默认 1.0E6
    tHomingTimeout      : TIME := T#60S;      // 回零总超时（Homing timeout），默认 T#60S，0=禁用
    bLimPos             : BOOL := FALSE;      // 正限位开关（Positive limit switch），TRUE=已压住
    bLimNeg             : BOOL := FALSE;      // 负限位开关（Negative limit switch），TRUE=已压住
    bHomeSw             : BOOL := FALSE;      // 原点开关（Home switch），TRUE=已压住
    bZeroPulse          : BOOL := FALSE;      // Z 相脉冲（Encoder zero pulse），捕获上升沿
    bTorqueLimitReached : BOOL := FALSE;      // 堵转阈值到达（Torque limit reached），由驱动层注入（接口无扭矩域，外部注入声明 R11 留档）
    bTrack              : BOOL := FALSE;      // 跟踪重同步（Track resync），TRUE 时中止序列回空闲（R19）
END_VAR
VAR_IN_OUT
    iAxis               : I_DL_MotionAxis;    // 轴接口引用（Axis reference），由上层注入实现块实例
END_VAR
VAR_OUTPUT
    bBusy               : BOOL := FALSE;      // 回零进行中（Homing busy）
    bDone               : BOOL := FALSE;      // 回零完成（Homing done），完成态保持至下次启动
    eStep               : E_DL_HomingStep := E_DL_HomingStep.eIdle; // 当前序列步（Current homing step），HMI 显示用
    uErrorId            : UDINT := 0;         // 末次事件码（Last error code），段位 16#0004_xxxx
END_VAR
VAR
    bInit               : BOOL := FALSE;      // 首扫标志（First-scan flag，R19 范式配套）
    bParamOk            : BOOL := FALSE;      // 参数门禁通过标志（Parameter gate pass flag），启动前逐拍重算
    bTmoEn              : BOOL := FALSE;      // 超时护栏使能（Timeout guard enable），tHomingTimeout > 0 时为 TRUE
    bTmoBreak           : BOOL := FALSE;      // 超时参数变更断拍标志（Timeout PT break flag，R14：变更后断输入一拍归零计时）
    tTmoLastRaw         : TIME := T#0S;       // 上一拍超时参数快照（Last timeout parameter snapshot，R14 配套）
    bAbortPend          : BOOL := FALSE;      // 中止挂起标志（Abort pending），受控停车完成后转已中止态
    bCmdSent            : BOOL := FALSE;      // 本步速度指令已发标志（Velocity command sent per step），换步自动复位
    bStopIssued         : BOOL := FALSE;      // 本步停止指令已发标志（Stop command sent per step），换步自动复位
    fDir                : REAL := 1.0;        // 回零方向系数（Direction factor），+1=正向 / -1=负向
    fVelHomEff          : REAL := 50.0;       // 生效快速逼近速度（Effective homing velocity）[mm/s]，恒正
    fVelCrpEff          : REAL := 2.0;        // 生效爬行速度（Effective creep velocity）[mm/s]，恒正
    fAccEff             : REAL := 1000.0;     // 生效加减速（Effective acceleration）[mm/s²]，防除零下限兜底
    fMaxTravelEff       : REAL := 1.0E6;      // 生效行程护栏（Effective travel guard）[mm]，非有限值兜底
    fVelApp             : REAL := 0.0;        // 逼近步带符号速度（Approach velocity signed）[mm/s]
    fVelRet             : REAL := 0.0;        // 限位回退步带符号速度（Limit retreat velocity signed）[mm/s]
    fVelCrpRev          : REAL := 0.0;        // 反向爬行带符号速度（Reverse creep velocity signed）[mm/s]
    fVelCrpFwd          : REAL := 0.0;        // 正向爬行带符号速度（Forward creep velocity signed）[mm/s]
    fStartPos           : REAL := 0.0;        // 启动时记录的起点位置（Start position snapshot）[mm]
    bLimWatch           : BOOL := FALSE;      // 当前模式监听的限位电平（Watched limit level），按 bDirNeg 选择
    eStepPrev           : E_DL_HomingStep := E_DL_HomingStep.eIdle; // 上一拍序列步（Previous step），换步复位步内标志
    rtrigStart          : R_TRIG;             // 启动指令上升沿（Rising edge of homing start）
    rtrigLimPos         : R_TRIG;             // 正限位上升沿（Rising edge of positive limit）
    rtrigLimNeg         : R_TRIG;             // 负限位上升沿（Rising edge of negative limit）
    rtrigHomeSw         : R_TRIG;             // 原点开关上升沿（Rising edge of home switch）
    rtrigZero           : R_TRIG;             // Z 相脉冲上升沿（Rising edge of zero pulse）
    rtrigTorque         : R_TRIG;             // 堵转信号上升沿（Rising edge of torque limit signal）
    ftrigLimPos         : F_TRIG;             // 正限位下降沿（Falling edge of positive limit）
    ftrigLimNeg         : F_TRIG;             // 负限位下降沿（Falling edge of negative limit）
    ftrigHomeSw         : F_TRIG;             // 原点开关下降沿（Falling edge of home switch）
    tonHome             : TON;                // 回零总超时定时器（Homing timeout timer）
END_VAR
VAR CONSTANT
    DL_HOM_INF_MAX      : REAL := 1.0E30;     // 有限值判定幅值上限（Finite-value magnitude bound）[mm]
    DL_HOM_EPS          : REAL := 1.0E-6;     // 浮点判零容差（Float zero tolerance）[mm]
    DL_HOM_VEL_FLOOR    : REAL := 1.0E-3;     // 速度/加速度参数下限（Velocity and acceleration floor）[mm/s 或 mm/s²]
END_VAR

METHOD IssueVel : BOOL
VAR_INPUT
    fV : REAL;                                   // 带符号速度指令（Signed velocity command）[mm/s]
END_VAR
IssueVel := iAxis.MoveVelocity(fV, fAccEff);     // 转发轴接口，受理结果即返回值
    END_METHOD

// 段 1｜沿检测与定时器无条件周期刷新（R7 红线，严禁置于分支内；实例入参先算成变量再喂实例）
rtrigStart(CLK := bCmdStart);
rtrigLimPos(CLK := bLimPos);      rtrigLimNeg(CLK := bLimNeg);
rtrigHomeSw(CLK := bHomeSw);
rtrigZero(CLK := bZeroPulse);     rtrigTorque(CLK := bTorqueLimitReached);
ftrigLimPos(CLK := bLimPos);      ftrigLimNeg(CLK := bLimNeg);
ftrigHomeSw(CLK := bHomeSw);
// R14：tHomingTimeout 语义参数变更时显式断输入一拍，使已计时归零
IF tHomingTimeout <> tTmoLastRaw THEN bTmoBreak := TRUE;  tTmoLastRaw := tHomingTimeout; END_IF
tonHome(IN := bBusy AND (NOT bTmoBreak), PT := tHomingTimeout);  // 回零总超时定时器（无条件刷新，R7）
bTmoBreak := FALSE;                              // 断拍标志本拍消费后复位

// 段 2｜接口引用有效性防御：未注入轴引用则直接退出（不产生误动作）
IF iAxis = 0 THEN
    bBusy := FALSE;
    RETURN;
END_IF

// 段 3｜R19 首扫/跟踪同步：判据唯一合法范式 IF bTrack OR (NOT bInit)
IF bTrack OR (NOT bInit) THEN
    IF bInit AND bBusy THEN
        iAxis.Stop();                            // 中途插入跟踪脉冲 → 受控停车
    END_IF
    eStep   := E_DL_HomingStep.eIdle;            // 中止序列回空闲（R19）
    bBusy   := FALSE;
    bAbortPend := FALSE;
    bCmdSent := FALSE;
    bStopIssued := FALSE;
    bInit   := TRUE;
END_IF

// 段 4｜参数防御与方向解析（公约 0.6/0.8）：非法参数仅封锁启动（信息级 0004_0106），不影响运行中扫描
fDir := 1.0;                                     // 方向系数默认正向 [1]
IF bDirNeg THEN fDir := -1.0; END_IF
bLimWatch := bLimPos;                            // 正向回零监听正限位
IF bDirNeg THEN bLimWatch := bLimNeg; END_IF     // 负向回零监听负限位
bParamOk := TRUE;
IF (fHomingVel <> fHomingVel) OR (fCreepVel <> fCreepVel) OR (fAcc <> fAcc)
   OR (fHomingVel <= DL_HOM_VEL_FLOOR) OR (fCreepVel <= DL_HOM_VEL_FLOOR)
   OR (fAcc <= DL_HOM_VEL_FLOOR)
   OR (fHomingVel > DL_HOM_INF_MAX) OR (fCreepVel > DL_HOM_INF_MAX)
   OR (fAcc > DL_HOM_INF_MAX) THEN
    bParamOk  := FALSE;                          // 速度/加速度非法或非有限值：拒绝启动
    fVelHomEff := 50.0;  fVelCrpEff := 2.0;  fAccEff := 1000.0;  // 安全兜底值，防运行中被改坏
ELSE
    fVelHomEff := fHomingVel;                    // 合法快速逼近速度直通 [mm/s]
    fVelCrpEff := fCreepVel;                     // 合法爬行速度直通 [mm/s]
    fAccEff    := fAcc;                          // 合法加减速直通 [mm/s²]
END_IF
IF (fMaxTravel <> fMaxTravel) OR (fMaxTravel <= DL_HOM_EPS) OR (fMaxTravel > DL_HOM_INF_MAX) THEN
    fMaxTravelEff := 1.0E6;                      // 行程护栏非法兜底 [mm]
    uErrorId := 16#0004_0106;                    // 信息级：参数兜底修复提示
ELSE
    fMaxTravelEff := fMaxTravel;                 // 合法行程护栏直通 [mm]
END_IF
bTmoEn := (tHomingTimeout > T#0MS);              // 超时 0=禁用护栏
fVelApp    := fDir * fVelCrpEff;                 // 逼近步默认爬行（Z 相/堵转模式）[mm/s]
IF (eMode = E_DL_HomingMode.eLimitSwitch) OR (eMode = E_DL_HomingMode.eHomeSwitch) THEN
    fVelApp := fDir * fVelHomEff;                // 限位/原点开关模式为快速逼近 [mm/s]
END_IF
fVelRet    := -fDir * fVelHomEff;                // 限位模式回退：全速反向 [mm/s]
fVelCrpRev := -fDir * fVelCrpEff;                // 原点开关模式反向爬行脱离 [mm/s]
fVelCrpFwd := fDir * fVelCrpEff;                 // 原点开关模式正向爬行再逼近 [mm/s]

// 段 5｜运行中全局护栏：轴故障 > 中止 > 超时 > 行程超限（优先级从高到低）
IF bBusy THEN
    IF iAxis.bError THEN
        eStep := E_DL_HomingStep.eFault;         // 轴故障：轴已自锁故障态，本块随之收口
        uErrorId := 16#0004_0212;
        bBusy := FALSE;
    ELSIF bCmdAbort THEN
        iAxis.Stop();                            // 中止：受控停车，停稳后转已中止态
        bAbortPend := TRUE;
        eStep := E_DL_HomingStep.eStopping;
    ELSIF bTmoEn AND tonHome.Q THEN
        iAxis.Stop();                            // 总超时：受控停车并锁存故障
        eStep := E_DL_HomingStep.eFault;
        uErrorId := 16#0004_0210;
        bBusy := FALSE;
    ELSIF ABS(iAxis.fPosition - fStartPos) > fMaxTravelEff THEN
        iAxis.Stop();                            // 行程超限：受控停车并锁存故障
        eStep := E_DL_HomingStep.eFault;
        uErrorId := 16#0004_0211;
        bBusy := FALSE;
    END_IF
END_IF

// 段 5.5｜终态重启借道（终审修复：eDone/eAborted/eFault 原为死态，启动沿被吞）：
//      三个终态收到启动上升沿 → 借道 eIdle，使下段 CASE 的 eIdle 门禁分支
//      同拍受理本次启动沿（边沿当拍仍有效，不吞沿、不双击）
IF rtrigStart.Q AND ((eStep = E_DL_HomingStep.eDone)
                  OR (eStep = E_DL_HomingStep.eAborted)
                  OR (eStep = E_DL_HomingStep.eFault)) THEN
    eStep := E_DL_HomingStep.eIdle;              // 终态重启：借道空闲态门禁（Restart from terminal state via idle gate）
END_IF

// 段 5.6｜换步检测：步号变化即复位步内指令标志（速度指令/停止指令各发一次）
IF eStep <> eStepPrev THEN
    bCmdSent := FALSE;
    bStopIssued := FALSE;
    eStepPrev := eStep;
END_IF

// 段 6｜回零序列状态机（ENUM + CASE + ELSE 兜底）
CASE eStep OF

    E_DL_HomingStep.eIdle:                       // 空闲态：等待启动门禁
        bBusy := FALSE;
        IF rtrigStart.Q THEN
            IF NOT bParamOk THEN
                uErrorId := 16#0004_0106;        // 参数门禁拒绝（信息级）
            ELSIF iAxis.eState <> E_DL_AxisState.eStandstill THEN
                uErrorId := 16#0004_0106;        // 轴不在待机态，拒绝启动（信息级）
            ELSIF (eMode = E_DL_HomingMode.eLimitSwitch) AND bLimWatch THEN
                uErrorId := 16#0004_0106;        // 可观测矛盾：启动时限位已压住
            ELSIF (eMode = E_DL_HomingMode.eHomeSwitch) AND bHomeSw THEN
                uErrorId := 16#0004_0106;        // 可观测矛盾：启动时原点开关已压住
            ELSE
                fStartPos := iAxis.fPosition;    // 记录行程护栏起点 [mm]
                bAbortPend := FALSE;
                bDone := FALSE;
                eStep := E_DL_HomingStep.eApproach;
            END_IF
        END_IF

    E_DL_HomingStep.eApproach:                   // 逼近态：按模式速度运行，监听参考事件
        bBusy := TRUE;
        IF NOT bCmdSent THEN
            IF IssueVel(fVelApp) THEN
                bCmdSent := TRUE;                // 速度指令受理，本步不再重发
            ELSE
                uErrorId := 16#0004_0213;        // 序列指令被轴拒绝（故障级）
                eStep := E_DL_HomingStep.eFault;
                bBusy := FALSE;
            END_IF
        ELSE
            CASE eMode OF
                E_DL_HomingMode.eLimitSwitch:    // 限位模式：监听所选限位上升沿
                    IF bDirNeg THEN
                        IF rtrigLimNeg.Q THEN bCmdSent := FALSE;  eStep := E_DL_HomingStep.eRetreat; END_IF
                    ELSE
                        IF rtrigLimPos.Q THEN bCmdSent := FALSE;  eStep := E_DL_HomingStep.eRetreat; END_IF
                    END_IF
                E_DL_HomingMode.eHomeSwitch:     // 原点开关模式：监听原点开关上升沿
                    IF rtrigHomeSw.Q THEN bCmdSent := FALSE;  eStep := E_DL_HomingStep.eRetreat; END_IF
                E_DL_HomingMode.eZeroPulse:      // Z 相模式：监听 Z 相上升沿
                    IF rtrigZero.Q THEN bCmdSent := FALSE;  eStep := E_DL_HomingStep.eCalibrate; END_IF
                E_DL_HomingMode.eTorqueBlock:    // 堵转模式：监听堵转信号上升沿
                    IF rtrigTorque.Q THEN bCmdSent := FALSE;  eStep := E_DL_HomingStep.eCalibrate; END_IF
                ELSE
                    uErrorId := 16#0004_0213;    // 非法模式兜底（故障级）
                    eStep := E_DL_HomingStep.eFault;
                    bBusy := FALSE;
            END_CASE
        END_IF

    E_DL_HomingStep.eRetreat:                    // 回退态：限位模式全速反向 / 原点开关模式停车后爬行脱离
        bBusy := TRUE;
        CASE eMode OF
            E_DL_HomingMode.eLimitSwitch:        // 限位模式：反向全速回退，监听限位下降沿确认脱离
                IF NOT bCmdSent THEN
                    IF IssueVel(fVelRet) THEN
                        bCmdSent := TRUE;
                    ELSE
                        uErrorId := 16#0004_0213;
                        eStep := E_DL_HomingStep.eFault;
                        bBusy := FALSE;
                    END_IF
                ELSIF bDirNeg THEN
                    IF ftrigLimNeg.Q THEN bCmdSent := FALSE;  eStep := E_DL_HomingStep.eReapproach; END_IF
                ELSE
                    IF ftrigLimPos.Q THEN bCmdSent := FALSE;  eStep := E_DL_HomingStep.eReapproach; END_IF
                END_IF
            E_DL_HomingMode.eHomeSwitch:         // 原点开关模式：先受控停车，停稳后反向爬行脱离
                IF NOT bStopIssued THEN
                    iAxis.Stop();                // 减速停（逼近沿触发）
                    bStopIssued := TRUE;
                ELSIF iAxis.eState = E_DL_AxisState.eStandstill THEN
                    IF NOT bCmdSent THEN
                        IF IssueVel(fVelCrpRev) THEN
                            bCmdSent := TRUE;
                        ELSE
                            uErrorId := 16#0004_0213;
                            eStep := E_DL_HomingStep.eFault;
                            bBusy := FALSE;
                        END_IF
                    ELSIF ftrigHomeSw.Q THEN     // 确认脱离原点开关（下降沿）
                        bCmdSent := FALSE;
                        eStep := E_DL_HomingStep.eReapproach;
                    END_IF
                END_IF
            ELSE
                uErrorId := 16#0004_0213;        // Z 相/堵转模式不应进入回退态：非法兜底
                eStep := E_DL_HomingStep.eFault;
                bBusy := FALSE;
        END_CASE

    E_DL_HomingStep.eReapproach:                 // 爬行再逼近态：监听参考事件二次触发
        bBusy := TRUE;
        IF NOT bCmdSent THEN
            IF IssueVel(fVelCrpFwd) THEN
                bCmdSent := TRUE;
            ELSE
                uErrorId := 16#0004_0213;
                eStep := E_DL_HomingStep.eFault;
                bBusy := FALSE;
            END_IF
        ELSE
            CASE eMode OF
                E_DL_HomingMode.eLimitSwitch:    // 限位模式：监听限位上升沿
                    IF bDirNeg THEN
                        IF rtrigLimNeg.Q THEN bCmdSent := FALSE;  eStep := E_DL_HomingStep.eCalibrate; END_IF
                    ELSE
                        IF rtrigLimPos.Q THEN bCmdSent := FALSE;  eStep := E_DL_HomingStep.eCalibrate; END_IF
                    END_IF
                E_DL_HomingMode.eHomeSwitch:     // 原点开关模式：监听原点开关上升沿
                    IF rtrigHomeSw.Q THEN bCmdSent := FALSE;  eStep := E_DL_HomingStep.eCalibrate; END_IF
                ELSE
                    uErrorId := 16#0004_0213;    // Z 相/堵转模式不应进入再逼近态：非法兜底
                    eStep := E_DL_HomingStep.eFault;
                    bBusy := FALSE;
            END_CASE
        END_IF

    E_DL_HomingStep.eCalibrate:                  // 标定态：本块仅收口（坐标系写入由上层联动 bDone）
        bBusy := TRUE;
        eStep := E_DL_HomingStep.eStopping;      // 转受控停车，停车指令由停车态统一发出

    E_DL_HomingStep.eStopping:                   // 受控停车态：等待轴停稳后收口
        bBusy := TRUE;
        IF NOT bStopIssued THEN
            iAxis.Stop();                        // 受控停车指令（MC_Stop 语义）
            bStopIssued := TRUE;
        ELSIF iAxis.eState = E_DL_AxisState.eStandstill THEN
            IF bAbortPend THEN
                eStep := E_DL_HomingStep.eAborted;  // 中止收口
                uErrorId := 16#0004_0212;
                bBusy := FALSE;
            ELSE
                eStep := E_DL_HomingStep.eDone;     // 正常标定收口
            END_IF
        END_IF

    E_DL_HomingStep.eDone:                       // 完成态：bDone 保持，启动沿经段 5.5 借道空闲态门禁重新回零
        bBusy := FALSE;
        bDone := TRUE;

    E_DL_HomingStep.eAborted:                    // 已中止态：启动沿经段 5.5 借道空闲态门禁重新回零
        bBusy := FALSE;

    E_DL_HomingStep.eFault:                      // 故障态：码已锁存，启动沿经段 5.5 借道空闲态门禁重试
        bBusy := FALSE;

    ELSE
        // 非法状态兜底（故障级）
        uErrorId := 16#0004_0213;
        eStep := E_DL_HomingStep.eFault;
        bBusy := FALSE;

END_CASE

// 段 7｜忙状态出口聚合（R20：量纲=布尔派生式，与序列步语义一致）
bBusy := (eStep = E_DL_HomingStep.eApproach) OR (eStep = E_DL_HomingStep.eRetreat)
      OR (eStep = E_DL_HomingStep.eReapproach) OR (eStep = E_DL_HomingStep.eCalibrate)
      OR (eStep = E_DL_HomingStep.eStopping);

(*-----------------------------------------------------------------------------
 * 方法实现（METHOD）：速度指令派发子过程，非阻塞，直接转发轴接口受理结果。
 *-----------------------------------------------------------------------------*)

END_FUNCTION_BLOCK

(* ---- FB_DL_DualEncoderDeviationWatch.st ---- *)
(*==============================================================================
 * 组件名称 (Component)  : FB_DL_DualEncoderDeviationWatch
 * 所属子库 (Sublibrary) : DL_Motion
 * 当前版本 (Version)    : 1.0.1
 * 兼容性   (Platform)   : CODESYS 3.5 / TwinCAT 3 / 汇川 InoProShop / 施耐德 Machine Expert
 *                         仅依赖 IEC 61131-3 标准库（TON / ABS / MAX），零厂商方言
 * 功能描述 (Function)   : 双编码器（电机侧 / 负载侧）位置与速度双反馈偏差监测：
 *                         ① 逐拍计算位置偏差 fDevPos 与速度偏差 fDevVel 的绝对值 [mm]/[mm/s]；
 *                         ② **启动屏蔽窗口**：bEnable 上升后 tBlank 时长内不产生预警 /
 *                            报警 / 停机请求，偏差仍照常计算便于投运观察；窗口由内部
 *                            锁存位 bBlankDone 一次性结束，bEnable 跌落即清锁存；
 *                         ③ **分级延时确认**：预警 tonWarn / 报警 tonAlarm / 停机 tonTrip
 *                            三个 TON 各自独立、无条件每周期刷新，延时到即按序晋级；
 *                         ④ **停机请求** bTripReq 锁存输出，解除路径唯一：
 *                            bReset 且偏差条件已消失（NOT bTripCond）；
 *                         ⑤ **编码器失效单独判定**：非有限值（NaN 自反 / Inf 阈值直比）
 *                            与单拍位置跳变（> fPosJumpMax）各自成码，任一编码器失效即
 *                            进 eFault，偏差不再用坏值重算（保持上一拍值并披露）。
 * 接口     (Interface)  : 输入 20 项（使能 / 复位 / 双侧位置速度 / 6 个分级阈值 /
 *                         跳变上限 / 4 个时间常数），输出 11 项（状态回执 / 双侧偏差 /
 *                         屏蔽窗回执 / 三级出口 / 编码器有效回执 / 有效性与故障码）。
 * 边界     (Boundary)   : ① 阈值做「≥ 1E-3 且 预警 ≤ 报警 ≤ 停机」递增序硬钳位，
 *                            钳位成立时置信息码 16#0004_1001（不置 bError）；
 *                         ② 屏蔽窗口只在 bEnable 上升沿开一次，不做周期重开；
 *                         ③ 编码器失效判定只覆盖「非有限」与「单拍跳变」两类，
 *                            不含断线 / 信号丢失（由上层硬件位在他件处理）；
 *                         ④ 本件只出停机**请求**位，不执行停机，执行由上层安全链完成；
 *                         ⑤ 零全局耦合（无 GVL / VAR_EXTERNAL / %I / %Q）。
 * 码表     (Codes)      : 本件占用 16#0004_1001 ~ 16#0004_100F 区间，实际使用 5 个：
 *                         1001 信息级 阈值钳位；1002 故障级 电机侧编码器失效；
 *                         1003 故障级 负载侧编码器失效；1004 信息级 偏差超预警；
 *                         1005 信息级 偏差超报警；1006 故障级 停机请求已锁存；
 *                         1008 故障级 非法状态兜底。信息级码永不置 bError。
 * 分工声明 (Scope)      : 与 FB_DL_AxisDualFeedbackGuard 分工：那件做闭环反馈切换与
 *                         位置给定仲裁；本件只做两侧偏差监测与分级保护请求。
 * 开源溯源 (Origin)     : 开源溯源：原创实现（无外部代码引入）
 * 红线自检 (Redline)    : R1 ✓ 零 GVL / VAR_EXTERNAL ｜ R2 ✓ 零 %I/%Q/%M
 *                         R3 ✓ 纯 IEC 61131-3 ｜ R4 ✓ 钳位 + 容差 1E-9 + 非有限双判
 *                         R5 ✓ 声明逐行同行双语注释 ｜ R6 ✓ 六态 ENUM + CASE + ELSE
 *                         R7 ✓ 四个 TON 无条件每周期调用
 * 修订历史 (Revision)   : 2026-11-23  v1.0.0  R77 首版
 *                         2026-11-23  v1.0.1  R77 闸修复（Inf 判据改阈值直比，修 Inf−Inf=NaN 致支路恒假）
 * 验收向量 (Acceptance) :
 *   V1 bEnable 上升、tBlank=2s、偏差 0 → 第 1 拍 eStateOut=eBlank，
 *      bBlankActive=TRUE，bWarn/bAlarm/bTripReq 全 FALSE；2s 后 eBlank → eMonitor。
 *   V2 屏蔽窗结束后位置偏差恒 1.5mm（预警 1.0 / 报警 2.0 / 停机 5.0）：
 *      tWarnDly 到后 bWarn=TRUE、eStateOut=eWarn、uErrorId=16#0004_1004、bError=FALSE。
 *   V3 位置偏差恒 6.0mm：tonTrip 到时 bTripReq=TRUE 且锁存，uErrorId=16#0004_1006、
 *      bError=TRUE；即使偏差回落到 0，bTripReq 仍 TRUE，直到 bReset 单拍。
 *   V4 电机侧 fPosMotor = NaN：本拍 bMotorEncValid=FALSE、eStateOut=eFault、
 *      uErrorId=16#0004_1002、fDevPos 保持上一拍值（不拿坏值重算）。
 *   V5 fPosLoad 单拍从 0 跳到 600.0（fPosJumpMax=500.0）：bLoadEncValid=FALSE、
 *      uErrorId=16#0004_1003；单拍后跳变锁存保持至 bReset。
 *============================================================================*)

(*-----------------------------------------------------------------------------
 * 调用示例 (Instance guide)：
 *   声明于调用方 FB 的 VAR 区：fbDew : FB_DL_DualEncoderDeviationWatch;
 *   每周期无条件调用：fbDew(bEnable := xRun, bReset := xReset,
 *                            fPosMotor := stAx.fActPosMotor, fPosLoad := stAx.fActPosLoad,
 *                            fVelMotor := stAx.fActVelMotor, fVelLoad := stAx.fActVelLoad);
 *   取用出口：IF fbDew.bTripReq THEN 触发上层安全链停止；诊断取 fbDew.uErrorId。
 *   调参指引：fDevWarnPos 取机械间隙的 1.5 倍，fDevAlarmPos 取 2 倍，
 *            fDevTripPos 取联轴器失效前的可辨认位差；tBlank 取启动加速段时长再加 20%。
 *----------------------------------------------------------------------------*)

(*-----------------------------------------------------------------------------
 * 枚举: E_DL_DewState（归属 DL_Motion，与 FB_DL_DualEncoderDeviationWatch 同文件）
 * 含义: 双编码器偏差监测状态机离散状态。eBlank 只覆盖启动屏蔽窗，eMonitor 为常规
 *       监测相，eWarn / eAlarm 为分级确认相，eFault 为编码器失效与非法状态兜底相。
 *----------------------------------------------------------------------------*)
TYPE E_DL_DewState :
(
    eInit    := 0,    // 首扫态：出口全部复位，等 bEnable 上升 / First scan: outputs reset, waiting for bEnable rise
    eBlank   := 10,   // 启动屏蔽窗态：只算偏差不报警，窗口结束转 eMonitor / Startup blanking: deviations computed, no alarms until window ends
    eMonitor := 20,   // 常规监测态：三级延时确认累积中 / Normal monitoring: three-level confirmation accumulating
    eWarn    := 30,   // 预警确认态：bWarn 置位，条件消失即退回 eMonitor / Warning state: bWarn set, falls back when condition clears
    eAlarm   := 40,   // 报警确认态：bAlarm 置位，停机延时继续累积 / Alarm state: bAlarm set, trip delay keeps accumulating
    eFault   := 99    // 故障兜底态：编码器失效或非法状态进入，锁存至 bReset / Fault fallback: encoder failure or illegal state, latched until bReset
);
END_TYPE

(*==============================================================================
 * 功能块: FB_DL_DualEncoderDeviationWatch
 * 调用约定: 每周期无条件调用一次；四个 TON 实例在段 3 无条件刷新，禁置于 CASE 内。
 * 屏蔽语义: bBlankActive = TRUE 期间，tonWarn / tonAlarm / tonTrip 的 IN 条件被
 *           bDevValid 与 NOT bBlankActive 共同门控，故延时不会在窗口内悄悄累积。
 *============================================================================*)
FUNCTION_BLOCK FB_DL_DualEncoderDeviationWatch
VAR_INPUT
    bEnable       : BOOL := FALSE;       // 监测使能，上升沿开启屏蔽窗，跌落清全部锁存 / Enable, rising edge opens blank window, falling clears all latches
    bReset        : BOOL := FALSE;       // 复位（电平有效），清停机锁存与跳变锁存 / Reset (level), clears trip latch and jump latches
    fPosMotor     : REAL := 0.0;         // 电机侧编码器位置反馈 [mm] / Motor-side encoder position feedback [mm]
    fPosLoad      : REAL := 0.0;         // 负载侧编码器位置反馈 [mm] / Load-side encoder position feedback [mm]
    fVelMotor     : REAL := 0.0;         // 电机侧编码器速度反馈 [mm/s] / Motor-side encoder velocity feedback [mm/s]
    fVelLoad      : REAL := 0.0;         // 负载侧编码器速度反馈 [mm/s] / Load-side encoder velocity feedback [mm/s]
    fDevWarnPos   : REAL := 1.0;         // 位置偏差预警阈值 [mm] / Position deviation warning threshold [mm]
    fDevAlarmPos  : REAL := 2.0;         // 位置偏差报警阈值 [mm] / Position deviation alarm threshold [mm]
    fDevTripPos   : REAL := 5.0;         // 位置偏差停机阈值 [mm] / Position deviation trip threshold [mm]
    fDevWarnVel   : REAL := 10.0;        // 速度偏差预警阈值 [mm/s] / Velocity deviation warning threshold [mm/s]
    fDevAlarmVel  : REAL := 20.0;        // 速度偏差报警阈值 [mm/s] / Velocity deviation alarm threshold [mm/s]
    fDevTripVel   : REAL := 50.0;        // 速度偏差停机阈值 [mm/s] / Velocity deviation trip threshold [mm/s]
    fPosJumpMax   : REAL := 500.0;       // 单拍位置跳变上限，超限判编码器失效 [mm] / Single-scan position jump limit, exceeding means encoder failure [mm]
    tBlank        : TIME := T#2S;        // 启动屏蔽窗口时长，T#0S = 不屏蔽直通 [s] / Startup blanking window, T#0S = no blanking [s]
    tWarnDly      : TIME := T#500MS;     // 预警确认延时 [s] / Warning confirmation delay [s]
    tAlarmDly     : TIME := T#300MS;     // 报警确认延时 [s] / Alarm confirmation delay [s]
    tTripDly      : TIME := T#2S;        // 停机请求确认延时 [s] / Trip request confirmation delay [s]
END_VAR
VAR_OUTPUT
    eStateOut     : E_DL_DewState;       // 状态机当前状态回执 [-] / Current state feedback of the state machine
    fDevPos       : REAL;                // 位置偏差绝对值，失效时保持上一拍 [mm] / Absolute position deviation, held on invalid [mm]
    fDevVel       : REAL;                // 速度偏差绝对值，失效时保持上一拍 [mm/s] / Absolute velocity deviation, held on invalid [mm/s]
    bBlankActive  : BOOL;                // 启动屏蔽窗口生效中，TRUE 期间不产生任何报警 / Blanking window active, no alarm during TRUE
    bWarn         : BOOL;                // 预警出口（信息级，不置 bError）/ Warning outlet, info level, keeps bError FALSE
    bAlarm        : BOOL;                // 报警出口（信息级，不置 bError）/ Alarm outlet, info level, keeps bError FALSE
    bTripReq      : BOOL;                // 停机请求出口（锁存，解除路径唯一：bReset 且条件消失）/ Trip request outlet, latched, cleared only by bReset with condition gone
    bMotorEncValid: BOOL;                // 电机侧编码器有效回执 / Motor-side encoder validity feedback
    bLoadEncValid : BOOL;                // 负载侧编码器有效回执 / Load-side encoder validity feedback
    bValid        : BOOL;                // 出口数据可信标志，失效相为 FALSE / Output data trustworthy flag, FALSE in invalid states
    bError        : BOOL;                // 故障级标志，与 uErrorId 严格联动 / Fault-level flag, strictly coupled with uErrorId
    uErrorId      : UDINT;               // 错误码，0 = 无码 / Error code, 0 = no code
END_VAR
VAR
    eState        : E_DL_DewState;       // 状态机内部当前状态 [-] / Internal current state
    tonBlank      : TON;                 // 启动屏蔽窗定时器（一次性，由锁存位终止）/ Startup blanking timer, one shot, terminated by latch
    tonWarn       : TON;                 // 预警确认延时定时器，无条件刷新 / Warning confirmation timer, refreshed unconditionally
    tonAlarm      : TON;                 // 报警确认延时定时器，无条件刷新 / Alarm confirmation timer, refreshed unconditionally
    tonTrip       : TON;                 // 停机请求确认延时定时器，无条件刷新 / Trip confirmation timer, refreshed unconditionally
    bBlankDone    : BOOL;                // 屏蔽窗结束锁存位，bEnable 跌落清零 / Blanking window finished latch, cleared when bEnable falls
    bBlankEn      : BOOL;                // 屏蔽功能是否启用（tBlank > 0）/ Blanking enabled flag, TRUE when tBlank > 0
    bBlankActiveI : BOOL;                // 内部屏蔽窗生效量，供 IN 条件引用 / Internal blanking active quantity used by IN conditions
    bWarnCond     : BOOL;                // 预警条件（已过域闸与屏蔽闸）/ Warning condition after domain and blanking gates
    bAlarmCond    : BOOL;                // 报警条件（已过域闸与屏蔽闸）/ Alarm condition after domain and blanking gates
    bTripCond     : BOOL;                // 停机条件（已过域闸与屏蔽闸，不受屏蔽窗影响以外）/ Trip condition after gates
    bDevValid     : BOOL;                // 本拍双侧编码器均有效、偏差可信 / Both encoders valid this scan, deviations trustworthy
    bMotorFinite  : BOOL;                // 电机侧反馈均为有限值 / Motor-side feedback values finite
    bLoadFinite   : BOOL;                // 负载侧反馈均为有限值 / Load-side feedback values finite
    bMotorNaN     : BOOL;                // 电机侧自反判 NaN 命中 / Motor-side NaN detected by self-comparison
    bMotorInf     : BOOL;                // 电机侧阈值直比判 Inf 命中 / Motor-side Infinity detected by direct threshold comparison
    bLoadNaN      : BOOL;                // 负载侧自反判 NaN 命中 / Load-side NaN detected by self-comparison
    bLoadInf      : BOOL;                // 负载侧阈值直比判 Inf 命中 / Load-side Infinity detected by direct threshold comparison
    bMotorJump    : BOOL;                // 电机侧单拍跳变锁存 / Motor-side single-scan jump latch
    bLoadJump     : BOOL;                // 负载侧单拍跳变锁存 / Load-side single-scan jump latch
    bHavePrev     : BOOL;                // 是否已有上一拍位置快照 / Previous position snapshot available
    fPrevPosMotor : REAL;                // 电机侧上一拍位置快照 [mm] / Motor-side previous position snapshot [mm]
    fPrevPosLoad  : REAL;                // 负载侧上一拍位置快照 [mm] / Load-side previous position snapshot [mm]
    bFaultLvl     : BOOL;                // 故障级标志内部量 / Internal fault-level flag
    fWarnPosEff   : REAL;                // 钳位后位置预警阈值 [mm] / Clamped position warning threshold [mm]
    fAlarmPosEff  : REAL;                // 钳位后位置报警阈值 [mm] / Clamped position alarm threshold [mm]
    fTripPosEff   : REAL;                // 钳位后位置停机阈值 [mm] / Clamped position trip threshold [mm]
    fWarnVelEff   : REAL;                // 钳位后速度预警阈值 [mm/s] / Clamped velocity warning threshold [mm/s]
    fAlarmVelEff  : REAL;                // 钳位后速度报警阈值 [mm/s] / Clamped velocity alarm threshold [mm/s]
    fTripVelEff   : REAL;                // 钳位后速度停机阈值 [mm/s] / Clamped velocity trip threshold [mm/s]
    fJumpEff      : REAL;                // 钳位后单拍跳变上限 [mm] / Clamped single-scan jump limit [mm]
    uInfoCode     : UDINT;               // 信息级码暂存（参数钳位等）/ Info-level code scratch, parameter clamping etc.
    bTripLatch    : BOOL;                // 停机请求锁存位 / Trip request latch
END_VAR
VAR CONSTANT
    DL_DEW_OK   : UDINT := 16#0000_0000; // 无码哨兵 / No-code sentinel
    DL_DEW_TOL  : REAL := 1.0E-3;        // 阈值下限硬钳位值，防零阈值抖动 [mm] / Threshold lower clamp preventing zero-threshold chatter
    DL_DEW_EPS  : REAL := 1.0E-9;        // 浮点比较容差（本件统一口径）/ Unified floating point comparison tolerance
    DL_DEW_ZERO : REAL := 0.0;           // 零基准哨兵 / Zero reference sentinel
    DL_DEW_HALF : REAL := 0.5;           // 中值系数（均值出口备用）/ Half factor for averaging outlet
    DL_DEW_RMAX : REAL := 3.4028235E38;  // 本机 REAL 可表示上限，Inf 阈值直比基准 [无量纲] / Locally representable REAL maximum, Inf threshold base
END_VAR

(*------------------------------------------------------------------------------
 * 段 0｜阈值域闸与钳位（不中断扫描）：强制递增序 预警 ≤ 报警 ≤ 停机，且均 ≥ 1E-3
 *      Threshold domain gate: enforce warning <= alarm <= trip and each >= 1E-3
 *      钳位一旦成立置信息码 16#0004_1001，不影响本拍监测能力（信息级不置 bError）
 *-----------------------------------------------------------------------------*)
uInfoCode    := DL_DEW_OK;                                  // 信息码预置无码 / Preset no info code
bFaultLvl    := FALSE;                                      // 故障级标志预置 / Preset fault-level flag FALSE

fWarnPosEff  := MAX(fDevWarnPos, DL_DEW_TOL);               // 位置预警阈值下限钳位 [mm] / Position warning lower clamp
fAlarmPosEff := MAX(fDevAlarmPos, fWarnPosEff);             // 位置报警阈值不低于预警 [mm] / Position alarm kept above warning
fTripPosEff  := MAX(fDevTripPos, fAlarmPosEff);             // 位置停机阈值不低于报警 [mm] / Position trip kept above alarm
fWarnVelEff  := MAX(fDevWarnVel, DL_DEW_TOL);               // 速度预警阈值下限钳位 [mm/s] / Velocity warning lower clamp
fAlarmVelEff := MAX(fDevAlarmVel, fWarnVelEff);             // 速度报警阈值不低于预警 [mm/s] / Velocity alarm kept above warning
fTripVelEff  := MAX(fDevTripVel, fAlarmVelEff);             // 速度停机阈值不低于报警 [mm/s] / Velocity trip kept above alarm
fJumpEff     := MAX(fPosJumpMax, DL_DEW_TOL);               // 跳变上限下限钳位 [mm] / Jump limit lower clamp

IF (ABS(fWarnPosEff - fDevWarnPos) > DL_DEW_EPS)
   OR (ABS(fAlarmPosEff - fDevAlarmPos) > DL_DEW_EPS)
   OR (ABS(fTripPosEff - fDevTripPos) > DL_DEW_EPS)
   OR (ABS(fWarnVelEff - fDevWarnVel) > DL_DEW_EPS)
   OR (ABS(fAlarmVelEff - fDevAlarmVel) > DL_DEW_EPS)
   OR (ABS(fTripVelEff - fDevTripVel) > DL_DEW_EPS)
   OR (ABS(fJumpEff - fPosJumpMax) > DL_DEW_EPS) THEN
    uInfoCode := 16#0004_1001;                              // 信息级：阈值越界已钳位 / Info: thresholds out of range, clamped
END_IF

(*------------------------------------------------------------------------------
 * 段 1｜编码器有效性判定：非有限（NaN 自反 / Inf 差自减）与单拍跳变分别成码
 *      Encoder validity: non-finite detection plus single-scan jump detection
 *      双判口径：NaN 用 x <> x 自反判；Inf 用「阈值直比」判（与 DL_DEW_RMAX 双侧比较），
 *      禁用 |x − x| 差自减口径——IEEE-754 下 Inf − Inf = NaN，任何与 NaN 的比较恒假，
 *      会让 +Inf 首拍绕过跳变闸（bHavePrev=FALSE）直接泄漏到 fDevPos 出口并误报编码器有效。
 *      NaN detection uses x <> x; Infinity uses direct threshold comparison against DL_DEW_RMAX.
 *      The former |x - x| test is banned: Inf - Inf = NaN makes every comparison FALSE.
 *-----------------------------------------------------------------------------*)
bMotorNaN := (fPosMotor <> fPosMotor) OR (fVelMotor <> fVelMotor);                            // 自反判 NaN / NaN by self-comparison
bMotorInf := (fPosMotor > DL_DEW_RMAX) OR (fPosMotor < -DL_DEW_RMAX)
          OR (fVelMotor > DL_DEW_RMAX) OR (fVelMotor < -DL_DEW_RMAX);                        // Inf 阈值直比 / Infinity by direct threshold comparison
bMotorFinite := NOT (bMotorNaN OR bMotorInf);                                                // 电机侧有限标志 / Motor side finite flag

bLoadNaN  := (fPosLoad <> fPosLoad) OR (fVelLoad <> fVelLoad);                               // 自反判 NaN / NaN by self-comparison
bLoadInf  := (fPosLoad > DL_DEW_RMAX) OR (fPosLoad < -DL_DEW_RMAX)
          OR (fVelLoad > DL_DEW_RMAX) OR (fVelLoad < -DL_DEW_RMAX);                           // Inf 阈值直比 / Infinity by direct threshold comparison
bLoadFinite := NOT (bLoadNaN OR bLoadInf);                                                   // 负载侧有限标志 / Load side finite flag

IF bHavePrev AND bMotorFinite THEN
    IF ABS(fPosMotor - fPrevPosMotor) > fJumpEff THEN
        bMotorJump := TRUE;                                 // 电机侧跳变锁存（bReset 解除）/ Motor jump latched, cleared by bReset
    END_IF
END_IF
IF bHavePrev AND bLoadFinite THEN
    IF ABS(fPosLoad - fPrevPosLoad) > fJumpEff THEN
        bLoadJump := TRUE;                                  // 负载侧跳变锁存（bReset 解除）/ Load jump latched, cleared by bReset
    END_IF
END_IF

IF bReset OR NOT bEnable THEN
    bMotorJump := FALSE;                                    // 跳变锁存解除路径之一：复位 / Jump latch clear path: reset
    bLoadJump  := FALSE;                                    // 跳变锁存解除路径之一：复位 / Jump latch clear path: reset
    bHavePrev  := FALSE;                                    // 位置快照作废，下次重新建立基准 / Drop snapshot, rebuild baseline next run
END_IF

bMotorEncValid := bMotorFinite AND NOT bMotorJump;          // 电机侧编码器有效回执 / Motor encoder validity
bLoadEncValid  := bLoadFinite AND NOT bLoadJump;            // 负载侧编码器有效回执 / Load encoder validity

IF bMotorFinite THEN
    fPrevPosMotor := fPosMotor;                             // 有限值才更新快照，坏值不得污染基准 / Update snapshot only on finite value
END_IF
IF bLoadFinite THEN
    fPrevPosLoad := fPosLoad;                               // 有限值才更新快照，坏值不得污染基准 / Update snapshot only on finite value
END_IF
IF bMotorFinite AND bLoadFinite THEN
    bHavePrev := TRUE;                                      // 双侧均有限才建立基准 / Baseline built only when both sides finite
END_IF

(*------------------------------------------------------------------------------
 * 段 2｜偏差计算：仅双侧有效时重算，任一失效保持上一拍值（不拿坏值重算）
 *      Deviation computation: recompute only when both sides valid, else hold
 *-----------------------------------------------------------------------------*)
bDevValid := bMotorEncValid AND bLoadEncValid;              // 偏差可信闸 / Deviation trustworthy gate
IF bDevValid THEN
    fDevPos := ABS(fPosMotor - fPosLoad);                   // 位置偏差绝对值 [mm] / Absolute position deviation [mm]
    fDevVel := ABS(fVelMotor - fVelLoad);                   // 速度偏差绝对值 [mm/s] / Absolute velocity deviation [mm/s]
END_IF

(*------------------------------------------------------------------------------
 * 段 3｜定时器组无条件刷新（红线 R7）+ 屏蔽窗口一次性锁存
 *      Unconditional timer refresh plus one-shot blanking window latch
 *      屏蔽窗口径：tBlank = 0 时 bBlankEn = FALSE，直通不屏蔽（防零时长除类退化）
 *-----------------------------------------------------------------------------*)
bBlankEn := tBlank > T#0S;                                  // 屏蔽功能启用判定，零时长直通 / Blanking enabled test, zero duration passes through

tonBlank(IN := bEnable AND bBlankEn AND NOT bBlankDone, PT := tBlank);   // 屏蔽窗计时，无条件调用 / Blanking timer, called unconditionally
IF NOT bEnable THEN
    bBlankDone := FALSE;                                    // 使能跌落清屏蔽锁存，下次启动重开 / Enable fall clears blanking latch
ELSIF tonBlank.Q THEN
    bBlankDone := TRUE;                                     // 窗口到时置锁存，IN 随之变 FALSE 停止计时 / Window elapsed, latch stops the timer
END_IF
bBlankActiveI := bEnable AND bBlankEn AND NOT bBlankDone AND NOT tonBlank.Q;   // 屏蔽窗生效内部量 / Internal blanking active quantity
bBlankActive  := bBlankActiveI;                             // 对外回执 / Outward feedback

bWarnCond  := bEnable AND bDevValid AND NOT bBlankActiveI
              AND ((fDevPos > fWarnPosEff) OR (fDevVel > fWarnVelEff));     // 预警条件（过域闸与屏蔽闸）/ Warning condition after gates
bAlarmCond := bEnable AND bDevValid AND NOT bBlankActiveI
              AND ((fDevPos > fAlarmPosEff) OR (fDevVel > fAlarmVelEff));   // 报警条件（过域闸与屏蔽闸）/ Alarm condition after gates
bTripCond  := bEnable AND bDevValid AND NOT bBlankActiveI
              AND ((fDevPos > fTripPosEff) OR (fDevVel > fTripVelEff));     // 停机条件（过域闸与屏蔽闸）/ Trip condition after gates

tonWarn(IN := bWarnCond, PT := tWarnDly);                   // 预警确认计时，无条件调用 / Warning delay timer, called unconditionally
tonAlarm(IN := bAlarmCond, PT := tAlarmDly);                // 报警确认计时，无条件调用 / Alarm delay timer, called unconditionally
tonTrip(IN := bTripCond, PT := tTripDly);                   // 停机确认计时，无条件调用 / Trip delay timer, called unconditionally

(*------------------------------------------------------------------------------
 * 段 4｜主状态机（红线 R6）：ENUM + CASE + ELSE 兜底
 *      Main state machine with enum, case coverage and ELSE interception
 *      入口约束：任何相迁入 eMonitor 前必须 bDevValid（数据可信），否则进 eFault
 *-----------------------------------------------------------------------------*)
CASE eState OF

    eInit:
        (* 首扫：出口全复位，等使能上升；屏蔽功能启用则先进 eBlank *)
        (* First scan: reset outlets, wait for enable, enter eBlank when blanking enabled *)
        bWarn  := FALSE;                                    // 预警出口复位 / Warning outlet reset
        bAlarm := FALSE;                                    // 报警出口复位 / Alarm outlet reset
        bValid := FALSE;                                    // 数据尚不可信 / Data not trustworthy yet
        IF bEnable THEN
            IF NOT bDevValid THEN
                eState := eFault;                           // 使能即失效：直接进故障相 / Invalid on enable, go to fault
            ELSIF bBlankEn THEN
                eState := eBlank;                           // 有屏蔽窗：先进 eBlank / Blanking enabled, enter eBlank
            ELSE
                eState := eMonitor;                         // 无屏蔽窗：直接进入监测 / No blanking, enter monitoring
            END_IF
        END_IF

    eBlank:
        (* 屏蔽窗：偏差照算但三级出口全压制，窗口结束转 eMonitor *)
        (* Blanking window: deviations computed but all alarm outlets suppressed *)
        bWarn  := FALSE;                                    // 窗口内不预警 / No warning inside the window
        bAlarm := FALSE;                                    // 窗口内不报警 / No alarm inside the window
        bValid := bDevValid;                                // 数据有效性照实回执 / Validity reported truthfully
        IF NOT bEnable THEN
            eState := eInit;                                // 使能跌落回首扫 / Enable drop returns to init
        ELSIF NOT bDevValid THEN
            eState := eFault;                               // 编码器失效立即进故障相 / Encoder failure goes to fault at once
        ELSIF NOT bBlankActiveI THEN
            eState := eMonitor;                             // 窗口结束（锁存位已置）进监测 / Window finished, enter monitoring
        END_IF

    eMonitor:
        (* 常规监测：三级延时按 停机 > 报警 > 预警 的优先级判定 *)
        (* Normal monitoring: trip outranks alarm which outranks warning *)
        bWarn  := FALSE;                                    // 监测相默认无预警 / No warning by default
        bAlarm := FALSE;                                    // 监测相默认无报警 / No alarm by default
        bValid := bDevValid;                                // 有效性照实回执 / Report validity truthfully
        IF NOT bEnable THEN
            eState := eInit;                                // 失能回首扫 / Disable returns to init
        ELSIF NOT bDevValid THEN
            eState := eFault;                               // 失效进故障相 / Invalid goes to fault
        ELSIF tonAlarm.Q THEN
            eState := eAlarm;                               // 报警延时到，直接进报警相 / Alarm delay elapsed, enter alarm
        ELSIF tonWarn.Q THEN
            eState := eWarn;                                // 预警延时到，进预警相 / Warning delay elapsed, enter warning
        END_IF

    eWarn:
        (* 预警相：退出条件 ≥2 条（报警沿晋级 / 预警条件消失退回）*)
        (* Warning state with two exit conditions: alarm rise or warning condition cleared *)
        bWarn  := TRUE;                                     // 预警出口置位 / Warning outlet set
        bAlarm := FALSE;                                    // 报警出口保持复位 / Alarm outlet stays reset
        bValid := bDevValid;                                // 有效性照实回执 / Report validity truthfully
        IF NOT bEnable THEN
            eState := eInit;                                // 失能回首扫 / Disable returns to init
        ELSIF NOT bDevValid THEN
            eState := eFault;                               // 失效进故障相 / Invalid goes to fault
        ELSIF tonAlarm.Q THEN
            eState := eAlarm;                               // 晋级报警 / Promote to alarm
        ELSIF NOT bWarnCond THEN
            eState := eMonitor;                             // 预警条件消失即退回监测 / Falls back when warning clears
        END_IF

    eAlarm:
        (* 报警相：停机延时继续累积；出口锁存由段 5 统一处理，本相不自清 *)
        (* Alarm state: trip delay keeps accumulating, latch handled in segment 5 *)
        bWarn  := TRUE;                                     // 报警相同时保持预警 / Warning held during alarm
        bAlarm := TRUE;                                     // 报警出口置位 / Alarm outlet set
        bValid := bDevValid;                                // 有效性照实回执 / Report validity truthfully
        IF NOT bEnable THEN
            eState := eInit;                                // 失能回首扫 / Disable returns to init
        ELSIF NOT bDevValid THEN
            eState := eFault;                               // 失效进故障相 / Invalid goes to fault
        ELSIF (NOT bAlarmCond) AND (NOT bTripLatch) THEN
            eState := eMonitor;                             // 报警条件消失且无停机锁存才退回 / Back only when alarm clears and no trip latch
        END_IF

    eFault:
        (* 故障兜底：出口全部压制，偏差保持上一拍；解除路径唯一：bReset 且双侧恢复有效 *)
        (* Fault fallback: outlets suppressed, deviations held, cleared only by bReset with both sides valid *)
        bWarn   := FALSE;                                   // 故障相不预警 / No warning in fault
        bAlarm  := FALSE;                                   // 故障相不报警 / No alarm in fault
        bValid  := FALSE;                                   // 数据不可信 / Data untrustworthy
        bFaultLvl := TRUE;                                  // 故障级标志置位 / Fault-level flag set
        IF bReset AND bMotorEncValid AND bLoadEncValid THEN
            eState := eMonitor;                             // 复位且恢复有效才解锁（跳变锁存已在段 1 清）/ Unlock only on reset with valid sides
        END_IF

    ELSE
        (* 非法状态拦截：任何未定义枚举值一律进故障相并置兜底码 *)
        (* Illegal state interception: undefined enum values go to fault with fallback code *)
        eState    := eFault;                                // 强制回故障相 / Force back to fault
        bWarn     := FALSE;                                 // 出口压制 / Outlet suppressed
        bAlarm    := FALSE;                                 // 出口压制 / Outlet suppressed
        bValid    := FALSE;                                 // 数据不可信 / Data untrustworthy
        bFaultLvl := TRUE;                                  // 故障级标志置位 / Fault-level flag set
        uInfoCode := 16#0004_1008;                          // 故障级：非法状态兜底 / Fault: illegal state fallback

END_CASE

(*------------------------------------------------------------------------------
 * 段 5｜停机请求锁存（置位唯一：tonTrip 到时；解除唯一：bReset 且 bTripCond 已消失）
 *      Trip request latch: set only on trip delay elapsed, cleared only by reset with condition gone
 *-----------------------------------------------------------------------------*)
IF bTripLatch THEN
    IF bReset AND (NOT bTripCond) THEN
        bTripLatch := FALSE;                                // 唯一解除路径：复位且偏差已回落 / Sole clear path: reset with deviation settled
    END_IF
ELSIF tonTrip.Q THEN
    bTripLatch := TRUE;                                     // 唯一置位路径：停机延时到 / Sole set path: trip delay elapsed
END_IF
bTripReq := bTripLatch;                                     // 对外锁存回放 / Latched replay to outlet

(*------------------------------------------------------------------------------
 * 段 6｜出口码统一映射（故障级锁存回放；信息级码永不置 bError，信息码仅当无更高优先级码时使用）
 *      Unified outlet code mapping: fault codes replayed, info codes never raise bError
 *-----------------------------------------------------------------------------*)
IF bTripLatch THEN
    uErrorId := 16#0004_1006;                               // 故障级：停机请求已锁存 / Fault: trip request latched
    bError   := TRUE;                                       // 故障级码配对置位 / Paired fault flag set
ELSIF NOT bMotorEncValid THEN
    uErrorId := 16#0004_1002;                               // 故障级：电机侧编码器失效 / Fault: motor-side encoder failed
    bError   := TRUE;                                       // 故障级码配对置位 / Paired fault flag set
ELSIF NOT bLoadEncValid THEN
    uErrorId := 16#0004_1003;                               // 故障级：负载侧编码器失效 / Fault: load-side encoder failed
    bError   := TRUE;                                       // 故障级码配对置位 / Paired fault flag set
ELSIF bAlarm THEN
    uErrorId := 16#0004_1005;                               // 信息级：偏差超报警阈值 / Info: deviation above alarm threshold
    bError   := FALSE;                                      // 信息级不置故障标志 / Info level never raises the fault flag
ELSIF bWarn THEN
    uErrorId := 16#0004_1004;                               // 信息级：偏差超预警阈值 / Info: deviation above warning threshold
    bError   := FALSE;                                      // 信息级不置故障标志 / Info level never raises the fault flag
ELSE
    uErrorId := uInfoCode;                                  // 参数钳位信息码或 0 / Parameter clamp info code or zero
    bError   := FALSE;                                      // 无故障级码即无故障 / No fault-level code means healthy
END_IF

eStateOut := eState;                                        // 状态回执（单一出口映射）/ State feedback through a single outlet
END_FUNCTION_BLOCK
